(* IEC 61131-3 sources: plcassist-cli/packages/volt-lsp-iec/test-corpus/bakon-nano/Device/Plc Logic/Application/Library Manager/L_MC1P_MotionControlBasic, 488 files *)

(* ---- L_MC1P_CONSTANTS.gvl ---- *)
VAR_GLOBAL
	GC_EPS : LREAL := 1E-10;
	GC_EPS_REAL : LREAL := 1E-06;
	GC_WUPDATEFILTER : WORD := 10;
	GC_WINSTANCENCHAR : WORD := 100;
	GC_WTRACEMAX : WORD := 100;
	GC_IMPLIZITCALLS : INT := 100;
	GC_MAXRETAINAXIS : INT := 256;
	GC_MAXAXISCOUNT : INT := 256;
	GC_ENCFILTERCYCLESMAX : INT := 100;
	GC_DWCHECKIDTAPPETREF : DWORD := 16#DC34;
	GC_SQRT2 : LREAL := 1.4142135623730951;
	GC_PI : LREAL := 3.1415926535897931;
	GC_REC_STATE : LWORD := SHL(1, 0);
	GC_REC_OPMODE : LWORD := SHL(1, 1);
	GC_REC_POS : LWORD := SHL(1, 2);
	GC_REC_VEL : LWORD := SHL(1, 3);
	GC_REC_TORQUE : LWORD := SHL(1, 4);
	GC_REC_ERRORID : LWORD := SHL(1, 5);
	GC_REC_FOLLERROR : LWORD := SHL(1, 6);
	GC_REC_STATELENZE : LWORD := SHL(1, 7);
	GC_REC_STATELENZE2 : LWORD := SHL(1, 8);
	GC_REC_TPSTATE1 : LWORD := SHL(1, 9);
	GC_REC_TP1POS : LWORD := SHL(1, 10);
	GC_REC_TP1NEG : LWORD := SHL(1, 11);
	GC_REC_TP2POS : LWORD := SHL(1, 12);
	GC_REC_TP2NEG : LWORD := SHL(1, 13);
	GC_REC_DIGIN : LWORD := SHL(1, 14);
	GC_REC_STATESM : LWORD := SHL(1, 15);
	GC_REC_VLACTVELOCITY : LWORD := SHL(1, 16);
	GC_REC_ENCPOS : LWORD := SHL(1, 17);
	GC_REC_ENCVEL : LWORD := SHL(1, 18);
	GC_REC_TP1POSTIME : LWORD := SHL(1, 19);
	GC_REC_TP1NEGTIME : LWORD := SHL(1, 20);
	GC_REC_TP2POSTIME : LWORD := SHL(1, 21);
	GC_REC_TP2NEGTIME : LWORD := SHL(1, 22);
	GC_REC_TPSTATE2 : LWORD := SHL(1, 23);
	GC_REC_TP3POS : LWORD := SHL(1, 24);
	GC_REC_TP3NEG : LWORD := SHL(1, 25);
	GC_REC_TP4POS : LWORD := SHL(1, 26);
	GC_REC_TP4NEG : LWORD := SHL(1, 27);
	GC_REC_TP3POSTIME : LWORD := SHL(1, 28);
	GC_REC_TP3NEGTIME : LWORD := SHL(1, 29);
	GC_REC_TP4POSTIME : LWORD := SHL(1, 30);
	GC_REC_TP4NEGTIME : LWORD := SHL(1, 31);
	GC_REC_SAFETYCTRL : LWORD := SHL(1, 32);
	GC_REC_SAFETYSTATE : LWORD := SHL(1, 33);
	GC_REC_SAFETYIOSTATE : LWORD := SHL(1, 34);
	GC_REC_ENCPOSTIMESTAMP : LWORD := SHL(1, 35);
	GC_REC_STATELENZEEXT : LWORD := SHL(1, 36);
	GC_REC_SPEEDERROR : LWORD := SHL(1, 37);
	GC_REC_POSVALUE1616 : LWORD := SHL(1, 38);
	GC_REC_CONTROLEFFORT : LWORD := SHL(1, 39);
	GC_REC_ACTPOSMOTORCIA402ADV : LWORD := SHL(1, 40);
	GC_REC_TEXTREFID : LWORD := SHL(1, 41);
	GC_REC_POSTIMESTAMP : LWORD := SHL(1, 42);
	GC_REC_MAXDATAINDEX : WORD := 43;
	GC_TRANS_CTRL : LWORD := SHL(1, 0);
	GC_TRANS_OPMODE : LWORD := SHL(1, 1);
	GC_TRANS_POS : LWORD := SHL(1, 2);
	GC_TRANS_VEL : LWORD := SHL(1, 3);
	GC_TRANS_TORQUE : LWORD := SHL(1, 4);
	GC_TRANS_TORQUELIMPOS : LWORD := SHL(1, 5);
	GC_TRANS_TORQUELIMNEG : LWORD := SHL(1, 6);
	GC_TRANS_SPEEDLIMUP : LWORD := SHL(1, 7);
	GC_TRANS_SPEEDLIMLOW : LWORD := SHL(1, 8);
	GC_TRANS_TPCTRL1 : LWORD := SHL(1, 9);
	GC_TRANS_POSOFFSET : LWORD := SHL(1, 10);
	GC_TRANS_VELOFFSET : LWORD := SHL(1, 11);
	GC_TRANS_TORQUEOFFSET : LWORD := SHL(1, 12);
	GC_TRANS_SPEEDCTRLINT : LWORD := SHL(1, 13);
	GC_TRANS_CTRLLENZE : LWORD := SHL(1, 14);
	GC_TRANS_VLTARGETVELOCITY : LWORD := SHL(1, 16);
	GC_TRANS_BRKOVRD : LWORD := SHL(1, 17);
	GC_TRANS_CTRLLENZE2 : LWORD := SHL(1, 18);
	GC_TRANS_CTRLLENZE3 : LWORD := SHL(1, 19);
	GC_TRANS_CTRLLENZE4 : LWORD := SHL(1, 20);
	GC_TRANS_TPCTRL2 : LWORD := SHL(1, 21);
	GC_TRANS_SAFEPOS : LWORD := SHL(1, 22);
	GC_TRANS_SAFEPOSSTATUS : LWORD := SHL(1, 23);
	GC_TRANS_SPEEDLIMITSLS : LWORD := SHL(1, 24);
	GC_TRANS_MAXDATAINDEX : WORD := 25;
	NODATAMEMORYAVAILABLE : WORD := WORD#16#1;
	MEMORYINVALID : WORD := WORD#16#2;
	MEMORYNOTINITIALIZED : WORD := WORD#16#4;
	NODATAAVAILABLE : WORD := WORD#16#8;
	NOMEMORYAVAILABLEFORAXIS : WORD := WORD#16#10;
	NOMEMORYINAXISARRAY : WORD := WORD#16#20;
	AXISGUIDCHANGED : WORD := WORD#16#40;
	C_SERIALNUMBER : UINT := 3;
	C_MANUFACTURER : UINT := 5;
	C_SOFTWAREREVISION : UINT := 9;
	C_HARDWAREREVISION : UINT := 10;
	C_DEVICECLASS : UINT := 11;
	C_PRODUCTCODE : UINT := 13;
	C_UPDATE : UINT := 99;
	C_CONNECTORTYPEMOTIONAXISOLD : UINT := 1279;
	C_CONNECTORTYPEMOTIONAXIS : UINT := 34279;
	C_CONNECTORTYPEENCODERIOSLICE : UINT := 33024;
END_VAR

(* ---- L_MC1P_INTERNAL.gvl ---- *)
VAR_GLOBAL
	DWDUMMY : DWORD;
	XAPPFIRSTRUN : BOOL := FALSE;
	PANYCONNECTOR : POINTER TO IoConfigConnector;
	LMAXISRETAINHANDLING : L_MC1P_AxisRetainMangaement;
	DWTIMESTAMPSIMU : DWORD;
	XTIMESTAMPUPDATED : BOOL;
	LMAXISMGMT : L_MC1P_AxisManagementFunction;
	CDIENUMSTARTVALUE : DINT := 50000;
END_VAR

(* ---- L_MC1P_IAXIS_REF_BRAKE.itf ---- *)
INTERFACE L_MC1P_IAXIS_REF_BRAKE
END_INTERFACE

METHOD GETACTVALUESBRAKE
END_METHOD

METHOD SWITCHONCONTROL
VAR_INPUT
	XSWITCHONREQUEST : BOOL;
END_VAR
VAR_OUTPUT
	XSWITCHON : BOOL;
END_VAR
VAR_IN_OUT
	AXIS : AXIS_REF;
END_VAR
END_METHOD

METHOD SWITCHEDONSTATUS
VAR_INPUT
	XSWITCHEDONREQUEST : BOOL;
END_VAR
VAR_OUTPUT
	XSWITCHEDON : BOOL;
END_VAR
VAR_IN_OUT
	AXIS : AXIS_REF;
END_VAR
END_METHOD

(* ---- L_MC1P_IAXIS_REF_MASTERVALUES.itf ---- *)
INTERFACE L_MC1P_IAXIS_REF_MASTERVALUES
END_INTERFACE

METHOD GETDIRECTION : WORD
VAR_INPUT
	VALUESOURCE : MC_SOURCE;
END_VAR
END_METHOD

METHOD GETMASTERERROR : BOOL
VAR_OUTPUT
	EERRORID : L_IE1P_Error;
END_VAR
END_METHOD

METHOD GETSTEADYSTATE : POINTER TO L_MC1P_SteadyState
END_METHOD

(* ---- L_MC1P_IAXIS_REF_POOL.itf ---- *)
INTERFACE L_MC1P_IAXIS_REF_POOL
END_INTERFACE

METHOD GETAXISFROMPOOL : POINTER TO AXIS_REF
VAR_INPUT
	WINDEX : WORD;
END_VAR
END_METHOD

(* ---- L_MC1P_IAXISCOMMMAND.itf ---- *)
INTERFACE L_MC1P_IAXISCOMMMAND
END_INTERFACE

METHOD ABORTING
END_METHOD

METHOD CALCSTATUS
VAR_IN_OUT
	AXIS : _AXIS_REF_REAL;
END_VAR
END_METHOD

METHOD EXECUTE
END_METHOD

METHOD MAIN
END_METHOD

METHOD RESETCOMMANDERRORSTATE : BOOL
VAR_IN_OUT
	AXIS : _AXIS_REF_REAL;
END_VAR
END_METHOD

METHOD RESETSTATUSPARAMETER
END_METHOD

METHOD SETINCTANCEINFO
VAR_INPUT
	PSINSTANCENAME : POINTER TO STRING;
	ERRORITFID : DWORD;
END_VAR
END_METHOD

METHOD UPDATEAXISPOINTER
VAR_INPUT
	PAXIS : POINTER TO AXIS_REF;
END_VAR
END_METHOD

METHOD UPDATECOMMANDINTERFACE
VAR_IN_OUT
	CMD : USINT;
END_VAR
END_METHOD

(* ---- L_MC1P_IAXISCOMMMAND_AUTOTUNING.itf ---- *)
INTERFACE L_MC1P_IAXISCOMMMAND_AUTOTUNING
END_INTERFACE

METHOD CALCPROFILEPARAMS
VAR_IN_OUT
	AXIS : AXIS_REF;
END_VAR
END_METHOD

METHOD UPDATEPARAINTERFACE
VAR_IN_OUT
	SCPAR : L_MC1P_AutotuningPara;
END_VAR
END_METHOD

(* ---- L_MC1P_IAXISEXTENSION.itf ---- *)
INTERFACE L_MC1P_IAXISEXTENSION
END_INTERFACE

METHOD SETBASICINITIALISATION
VAR_INPUT
	ITFGENERICCONFIG : L_MC1P_IGenericAxisConfiguration;
END_VAR
VAR_IN_OUT
	AXIS : _AXIS_REF_REAL;
END_VAR
END_METHOD

(* ---- L_MC1P_IAXISSIMCALLSINGLESTEPS.itf ---- *)
INTERFACE L_MC1P_IAXISSIMCALLSINGLESTEPS
END_INTERFACE

METHOD SIMFINISH : BOOL
VAR_INPUT
	AXISID : INT;
	ITFMECHANICSIMULATION : L_MC1P_IMechanicSimulation;
END_VAR
VAR_IN_OUT
	AXIS : _AXIS_REF_REAL;
END_VAR
END_METHOD

METHOD SIMINSIDELOOP : BOOL
VAR_INPUT
	AXISID : INT;
	ISYSTEMSIMCOUNTER : INT;
	ITFMECHANICSIMULATION : L_MC1P_IMechanicSimulation;
END_VAR
END_METHOD

METHOD SIMPREPARE : BOOL
VAR_INPUT
	AXISID : INT;
	ITFMECHANICSIMULATION : L_MC1P_IMechanicSimulation;
END_VAR
VAR_IN_OUT
	AXIS : _AXIS_REF_REAL;
END_VAR
END_METHOD

(* ---- L_MC1P_IAXISSIMULATIONINTERFACE.itf ---- *)
INTERFACE L_MC1P_IAXISSIMULATIONINTERFACE
END_INTERFACE

METHOD ACTIVATESIMULATION
VAR_IN_OUT
	AXIS : _AXIS_REF_REAL;
END_VAR
END_METHOD

METHOD CALCULATEINPUTDATA
VAR_INPUT
	ITFKINSIM : L_MC1P_IKinematicSimulation;
END_VAR
VAR_IN_OUT
	AXIS : _AXIS_REF_REAL;
END_VAR
END_METHOD

METHOD CALCULATEOUTPUTDATA
VAR_INPUT
	ITFKINSIM : L_MC1P_IKinematicSimulation;
END_VAR
VAR_IN_OUT
	AXIS : _AXIS_REF_REAL;
END_VAR
END_METHOD

METHOD DISABLESIMULATION
VAR_IN_OUT
	AXIS : _AXIS_REF_REAL;
END_VAR
END_METHOD

(* ---- L_MC1P_ICOMMMUNICATIONSIMULATION.itf ---- *)
INTERFACE L_MC1P_ICOMMMUNICATIONSIMULATION
END_INTERFACE

METHOD GETCOMMSTATE : L_DCO_CommState
VAR_INPUT
	PAXISCOMM : POINTER TO _AXIS_REF_COM;
END_VAR
END_METHOD

METHOD PARREAD
VAR_INPUT
	WIDX : DWORD;
END_VAR
END_METHOD

METHOD PARREAD_GETOUTPUT
VAR_INPUT
	WIDX : DWORD;
END_VAR
VAR_OUTPUT
	SZDATAREAD : CAA_SIZE;
	XDONE : BOOL;
	XERROR : BOOL;
	WERROR : WORD;
END_VAR
END_METHOD

METHOD PARREAD_SETINPUT
VAR_INPUT
	WIDX : DWORD;
	XEXECUTE : BOOL;
	WINDEX : WORD;
	BYSUBINDEX : BYTE;
	PBUFFER : POINTER TO BYTE;
	SZSIZE : UDINT;
	UDITIMEOUT : UDINT;
	XSLOTB : BOOL;
END_VAR
END_METHOD

METHOD PARWRITE
VAR_INPUT
	WIDX : DWORD;
END_VAR
END_METHOD

METHOD PARWRITE_GETOUTPUT
VAR_INPUT
	WIDX : DWORD;
END_VAR
VAR_OUTPUT
	XDONE : BOOL;
	XERROR : BOOL;
	WERROR : WORD;
END_VAR
END_METHOD

METHOD PARWRITE_SETINPUT
VAR_INPUT
	WIDX : DWORD;
	XEXECUTE : BOOL;
	WINDEX : WORD;
	BYSUBINDEX : BYTE;
	PBUFFER : POINTER TO BYTE;
	SZSIZE : UDINT;
	UDITIMEOUT : UDINT;
	XSLOTB : BOOL;
END_VAR
END_METHOD

METHOD RESTARTMASTER
VAR_INPUT
	XEXECUTE : BOOL;
	PAXIS : POINTER TO _AXIS_REF_COM;
END_VAR
VAR_OUTPUT
	XDONE : BOOL;
	XERROR : BOOL;
	XBUSY : BOOL;
	DWERROR : DWORD;
END_VAR
END_METHOD

(* ---- L_MC1P_ICOMMUNICATION.itf ---- *)
INTERFACE L_MC1P_ICOMMUNICATION
END_INTERFACE

METHOD FORWARDERROR
VAR_INPUT
	XENABLE : BOOL;
	XWARNING : BOOL;
	XERROR : BOOL;
	WERRORID : WORD;
	WTEXTREFID : WORD;
	XRESETERROR : BOOL := FALSE;
	AXISMODULEHANDLER : L_IMHP_IModuleHandler;
END_VAR
END_METHOD

METHOD GETCOMMPARAMETER
VAR_INPUT
	PCONNECTOR : POINTER TO IoConfigConnector;
END_VAR
VAR_OUTPUT
	PSLAVECONNECTOR : POINTER TO IoStandard.IoConfigConnector;
	UINETID : UINT;
	UIDEVICEID : UINT;
	XSENDFRAMEATTASKSTART : BOOL;
	UDIPRODUCTCODE : DWORD;
	PMASTERCONNECTOR : POINTER TO IoStandard.IoConfigConnector;
END_VAR
END_METHOD

METHOD GETCOMMSTATE : L_DCO_CommState
VAR_INPUT
	PAXISCOMM : POINTER TO _AXIS_REF_COM;
END_VAR
END_METHOD

METHOD GETPDINEQPDOUT : BOOL
END_METHOD

METHOD PARREAD
VAR_INPUT
	WIDX : DWORD;
END_VAR
END_METHOD

METHOD PARREAD_GETOUTPUT
VAR_INPUT
	WIDX : DWORD;
END_VAR
VAR_OUTPUT
	SZDATAREAD : CAA_SIZE;
	XDONE : BOOL;
	XERROR : BOOL;
	WERROR : WORD;
END_VAR
END_METHOD

METHOD PARREAD_SETINPUT
VAR_INPUT
	WIDX : DWORD;
	XEXECUTE : BOOL;
	WINDEX : WORD;
	BYSUBINDEX : BYTE;
	PBUFFER : POINTER TO BYTE;
	SZSIZE : UDINT;
	UDITIMEOUT : UDINT;
END_VAR
END_METHOD

METHOD PARWRITE
VAR_INPUT
	WIDX : DWORD;
END_VAR
END_METHOD

METHOD PARWRITE_GETOUTPUT
VAR_INPUT
	WIDX : DWORD;
END_VAR
VAR_OUTPUT
	XDONE : BOOL;
	XERROR : BOOL;
	WERROR : WORD;
END_VAR
END_METHOD

METHOD PARWRITE_SETINPUT
VAR_INPUT
	WIDX : DWORD;
	XEXECUTE : BOOL;
	WINDEX : WORD;
	BYSUBINDEX : BYTE;
	PBUFFER : POINTER TO BYTE;
	SZSIZE : UDINT;
	UDITIMEOUT : UDINT;
END_VAR
END_METHOD

METHOD RESET
END_METHOD

METHOD RESTARTMASTER
VAR_INPUT
	XEXECUTE : BOOL;
	PAXIS : POINTER TO _AXIS_REF_COM;
END_VAR
VAR_OUTPUT
	XDONE : BOOL;
	XERROR : BOOL;
	XBUSY : BOOL;
	DWERROR : DWORD;
END_VAR
END_METHOD

METHOD SETBASICINITIALISATION
VAR_IN_OUT
	AXIS : _AXIS_REF_REAL;
END_VAR
END_METHOD

METHOD SETCOMPONENTINFO
VAR_INPUT
	DATASELECTION : WORD;
	SDATA : STRING;
END_VAR
END_METHOD

(* ---- L_MC1P_ICOMPENSATIONINTERFACE.itf ---- *)
INTERFACE L_MC1P_ICOMPENSATIONINTERFACE
END_INTERFACE

METHOD GETOFFSETVALUES
VAR_OUTPUT
	LROFFSETPOS : LREAL;
	LROFFSETVEL : LREAL;
	LROFFSETACC : LREAL;
END_VAR
END_METHOD

(* ---- L_MC1P_ICONFIGUREDRIVE.itf ---- *)
INTERFACE L_MC1P_ICONFIGUREDRIVE
END_INTERFACE

METHOD DOFUNCTION : BOOL
VAR_INPUT
	XEXECUTE : BOOL;
	WOFFSET : WORD;
END_VAR
VAR_OUTPUT
	XDONE : BOOL;
	XERROR : BOOL;
	XBUSY : BOOL;
	EERRORID : WORD;
END_VAR
VAR_IN_OUT
	AXIS : _AXIS_REF_REAL;
END_VAR
END_METHOD

METHOD GETADDITIONALCONFIGINFO : POINTER TO L_MC1P_AdditionalConfigInfo
END_METHOD

METHOD GETINSTANCE : POINTER TO BYTE
END_METHOD

METHOD RESET : BOOL
END_METHOD

(* ---- L_MC1P_ICONTROLLERADAPTION.itf ---- *)
INTERFACE L_MC1P_ICONTROLLERADAPTION
END_INTERFACE

METHOD CALCADAPTIONCURVE : LREAL
VAR_INPUT
	LRSETVEL : LREAL;
END_VAR
VAR_IN_OUT
	AXIS : _AXIS_REF_REAL;
END_VAR
END_METHOD

(* ---- L_MC1P_ICONTROLLERINTERFACE.itf ---- *)
INTERFACE L_MC1P_ICONTROLLERINTERFACE
END_INTERFACE

METHOD CALCCONTROLLER
VAR_INPUT
	LRSETPOSITION : LREAL;
	LRSETVELOCITY : LREAL;
	LRSETACCELERATION : LREAL;
	LRSETTORQUE : LREAL;
	LRSETJERK : LREAL;
	LRACTPOSITIONIN : LREAL;
	LRACTVELOCITYIN : LREAL;
	LRACTACCELERATIONIN : LREAL;
	LRACTTORQUEIN : LREAL;
END_VAR
VAR_OUTPUT
	LRSETPOSITIONOUT : LREAL;
	LRSETVELOCITYOUT : LREAL;
	LRSETACCELERATIONOUT : LREAL;
	LRSETTORQUEOUT : LREAL;
END_VAR
VAR_IN_OUT
	AXIS : _AXIS_REF_REAL;
END_VAR
END_METHOD

(* ---- L_MC1P_IDRIVESCALING.itf ---- *)
INTERFACE L_MC1P_IDRIVESCALING
END_INTERFACE

METHOD CALCACCFACTOR : BOOL
VAR_OUTPUT
	LRSCALEUNITTOACC : LREAL;
	LRSCALEACCTOUNIT : LREAL;
END_VAR
VAR_IN_OUT
	AXIS : _AXIS_REF_REAL;
END_VAR
END_METHOD

METHOD CALCSPEEDFACTOR : BOOL
VAR_OUTPUT
	LRSCALEUNITTOSPEED : LREAL;
	LRSCALESPEEDTOUNIT : LREAL;
END_VAR
VAR_IN_OUT
	AXIS : _AXIS_REF_REAL;
END_VAR
END_METHOD

METHOD CALCTORQUEFACTOR : BOOL
VAR_OUTPUT
	LRSCALETORQUETONORM : LREAL;
	LRSCALETORQUETONORM2 : LREAL;
	LRSCALENORMTOTORQUE : LREAL;
END_VAR
VAR_IN_OUT
	AXIS : _AXIS_REF_REAL;
END_VAR
END_METHOD

METHOD CHECKVALIDPOSRESOLUTION : BOOL
VAR_INPUT
	DWPOSRESOLUTION : DWORD;
END_VAR
END_METHOD

METHOD GETDEFAULTTORQUE : LREAL
VAR_INPUT
	LRREFTORQUE : LREAL;
END_VAR
END_METHOD

METHOD POSDIFFTOSPEEDINC : DINT
VAR_INPUT
	DIPOSDIFF : DINT := 0;
	DWFACTOR : DWORD := 1000;
END_VAR
VAR_IN_OUT
	AXIS : _AXIS_REF_REAL;
END_VAR
END_METHOD

METHOD SPEEDTOPOSDIFFINC : DINT
VAR_INPUT
	DISPEED : DINT := 0;
	DWFACTOR : DWORD := 1000;
END_VAR
VAR_IN_OUT
	AXIS : _AXIS_REF_REAL;
	DIRES : DINT;
END_VAR
END_METHOD

(* ---- L_MC1P_IDRIVESPECIFICIMPLBASE.itf ---- *)
INTERFACE L_MC1P_IDRIVESPECIFICIMPLBASE
END_INTERFACE

METHOD CALCAFTERREADINPUTS
VAR_IN_OUT
	AXIS : _AXIS_REF_REAL;
END_VAR
END_METHOD

METHOD CALCBEFOREREADINPUTS
VAR_IN_OUT
	AXIS : _AXIS_REF_REAL;
END_VAR
END_METHOD

METHOD CALCBEFOREWRITEOUTPUTS
VAR_IN_OUT
	AXIS : _AXIS_REF_REAL;
END_VAR
END_METHOD

METHOD CHECKAVAILABLECONTROLMODE : BOOL
VAR_IN_OUT
	AXIS : _AXIS_REF_REAL;
	POSCTRLDRIVEAVAILABLE : L_IE1P_Error;
	POSCTRLPLCAVAILABLE : L_IE1P_Error;
	SPEEDCTRLDRIVEAVAILABLE : L_IE1P_Error;
	TORQUECTRLDRIVE : L_IE1P_Error;
END_VAR
END_METHOD

METHOD CHECKRESETHOMEPOS
VAR_INPUT
	WFDBSTATUSWORD : WORD;
END_VAR
VAR_IN_OUT
	AXIS : _AXIS_REF_REAL;
END_VAR
END_METHOD

METHOD CHECKSAFETYOPTIONAVAILABLE : BOOL
VAR_INPUT
	DWPRODUCTCODE : DWORD;
END_VAR
END_METHOD

METHOD COLLECTDRIVESTATE : BOOL
VAR_IN_OUT
	AXIS : _AXIS_REF_REAL;
	SCSTATEINFO : L_MC1P_DriveStateCollection;
END_VAR
END_METHOD

METHOD CONTROLDRIVE : BOOL
VAR_INPUT
	XENABLE : BOOL;
END_VAR
VAR_IN_OUT
	AXIS : _AXIS_REF_REAL;
END_VAR
END_METHOD

METHOD DRIVECONFIGDATA
VAR_INPUT
	PCONFIGINFO : POINTER TO L_MC1P_AdditionalConfigInfo;
END_VAR
VAR_IN_OUT
	AXIS : _AXIS_REF_REAL;
END_VAR
END_METHOD

METHOD DRIVEFAULTSTATUS : BOOL
VAR_IN_OUT
	AXIS : _AXIS_REF_REAL;
	SCSTATEINFO : L_MC1P_DriveStateCollection;
END_VAR
END_METHOD

METHOD GETBRAKE : POINTER TO L_MC1P_BrakeControlBase
VAR_IN_OUT
	AXIS : _AXIS_REF_REAL;
END_VAR
END_METHOD

METHOD GETBRAKESERVICE : POINTER TO L_MC1P_BrakeService
VAR_IN_OUT
	AXIS : _AXIS_REF_REAL;
END_VAR
END_METHOD

METHOD GETCAUSEOFCINH : WORD
VAR_IN_OUT
	AXIS : _AXIS_REF_REAL;
END_VAR
END_METHOD

METHOD GETFDBSTATUSWORD : WORD
VAR_IN_OUT
	AXIS : _AXIS_REF_REAL;
END_VAR
END_METHOD

METHOD GETIECADRESS : BOOL
VAR_IN_OUT
	AXIS : _AXIS_REF_REAL;
	M_PPDOINFOCONNECTOR : POINTER TO IoConfigConnector;
	ATRANSELEMENT : ARRAY [1.._AXIS_REF_REAL.c_wMaxTransElem] OF L_MC1P_MappedElement;
	WTRANSELEMENTS : WORD;
	LWTRANSDATA : LWORD;
	LWRECDATA : LWORD;
	WRECEIVEELEMENTS : WORD;
	ARECEIVEELEMENT : ARRAY [1.._AXIS_REF_REAL.c_wMaxRecElem] OF L_MC1P_MappedElement;
END_VAR
END_METHOD

METHOD GETOPTIONALACTVEL : BOOL
VAR_IN_OUT
	LRVEL : LREAL;
END_VAR
END_METHOD

METHOD GETRECEIVEDATAIMPL : DWORD
VAR_INPUT
	LWMASK : LWORD;
END_VAR
VAR_IN_OUT
	AXIS : _AXIS_REF_REAL;
END_VAR
END_METHOD

METHOD GETSTATUSWORDS
VAR_OUTPUT
	STATUSWORD1 : WORD;
	STATUSWORD2 : WORD;
	STATUSWORD3 : WORD;
	STATUSWORD4 : WORD;
END_VAR
VAR_IN_OUT
	AXIS : _AXIS_REF_REAL;
END_VAR
END_METHOD

METHOD GETTRANSMITDATAIMPL : DWORD
VAR_INPUT
	LWMASK : LWORD;
END_VAR
VAR_IN_OUT
	AXIS : _AXIS_REF_REAL;
END_VAR
END_METHOD

METHOD GETTRANSMITDATALREALIMPL : LREAL
VAR_INPUT
	LWMASK : LWORD;
END_VAR
VAR_IN_OUT
	AXIS : _AXIS_REF_REAL;
END_VAR
END_METHOD

METHOD HOMECONFIG : BOOL
VAR_INPUT
	LRPOSITION : LREAL;
END_VAR
VAR_OUTPUT
	WINDEX : WORD;
	BYSUBINDEX : BYTE;
	BYNROFBYTE : BYTE;
	DWDATA : DWORD;
	XWRITEPARAM : BOOL;
	XDONE : BOOL;
	XERROR : BOOL;
END_VAR
VAR_IN_OUT
	AXIS : _AXIS_REF_REAL;
	SCHOMEDATA : L_MC1P_HomeParameter;
	WSTEP : WORD;
END_VAR
END_METHOD

METHOD HOMEPOSPERMANENTSETACTIVE : BOOL
VAR_IN_OUT
	AXIS : _AXIS_REF_REAL;
END_VAR
END_METHOD

METHOD RECEIVEPARAMETER
VAR_INPUT
	WPARAMETER : WORD;
	PADRESS : POINTER TO BYTE;
	WSIZE : WORD;
END_VAR
VAR_IN_OUT
	AXIS : _AXIS_REF_REAL;
END_VAR
END_METHOD

METHOD RECEIVEPARAMETERCALC
VAR_IN_OUT
	AXIS : _AXIS_REF_REAL;
	DATA : ARRAY [1..L_MC1P_Constants.gc_Rec_MaxDataIndex] OF POINTER TO L_MC1P_MappedElement;
END_VAR
END_METHOD

METHOD RESETDRIVECONTROL
VAR_INPUT
	XRESETDRIVEERROR : BOOL;
END_VAR
END_METHOD

METHOD RESTOREADDITIONALRETAINDATA
VAR_INPUT
	PDATA : POINTER TO L_MC1P_uRetainData;
END_VAR
END_METHOD

METHOD SETAXISPROPERTIES
VAR_IN_OUT
	AXIS : _AXIS_REF_REAL;
	AXISPROPERTIES : L_MC1P_AxisProperties;
END_VAR
END_METHOD

METHOD SETAXISSTATUSWORD
VAR_IN_OUT
	AXIS : _AXIS_REF_REAL;
	DWAXISSTATUS : DWORD;
END_VAR
END_METHOD

METHOD SETBASICINITIALISATION
VAR_IN_OUT
	AXIS : _AXIS_REF_REAL;
END_VAR
END_METHOD

METHOD SETCONTROLWORDS
VAR_INPUT
	CONTROLWORD1 : WORD;
	CONTROLWORD2 : WORD;
	CONTROLWORD3 : WORD;
	CONTROLWORD4 : WORD;
END_VAR
VAR_IN_OUT
	AXIS : _AXIS_REF_REAL;
END_VAR
END_METHOD

METHOD SETDCBRAKE
VAR_INPUT
	XSETDCBRAKE : BOOL;
END_VAR
VAR_OUTPUT
	XDCBRAKEACTIVE : BOOL;
END_VAR
VAR_IN_OUT
	AXIS : _AXIS_REF_REAL;
END_VAR
END_METHOD

METHOD SETDRIVECONFIGINIT
VAR_IN_OUT
	AXIS : _AXIS_REF_REAL;
END_VAR
END_METHOD

METHOD SETSPEEDCTRLLIMITATION : BOOL
VAR_INPUT
	XLIMIT : BOOL;
END_VAR
VAR_IN_OUT
	AXIS : _AXIS_REF_REAL;
END_VAR
END_METHOD

METHOD SETSPEEDCTRLLOADVALUE
VAR_INPUT
	XLOAD : BOOL;
	LRVALUE : LREAL;
END_VAR
VAR_IN_OUT
	AXIS : _AXIS_REF_REAL;
END_VAR
END_METHOD

METHOD STOREADDITIONALRETAINDATA
VAR_INPUT
	PDATA : POINTER TO L_MC1P_uRetainData;
END_VAR
END_METHOD

METHOD TRANSMITPARAMETER
VAR_INPUT
	WPARAMETER : WORD;
	PADRESS : POINTER TO BYTE;
	WSIZE : WORD;
END_VAR
VAR_IN_OUT
	AXIS : _AXIS_REF_REAL;
END_VAR
END_METHOD

METHOD TRANSMITPARAMETERCALC
VAR_IN_OUT
	AXIS : _AXIS_REF_REAL;
	DATA : ARRAY [1..L_MC1P_Constants.gc_Trans_MaxDataIndex] OF POINTER TO L_MC1P_MappedElement;
END_VAR
END_METHOD

METHOD UPDATEMAPPING
VAR_INPUT
	PTASKMAPLIST : POINTER TO IoStandard.IoConfigTaskMap;
	NCOUNT : DINT;
	PPDOINFOCONNECTOR : POINTER TO IoConfigConnector;
END_VAR
VAR_IN_OUT
	AXIS : _AXIS_REF_REAL;
END_VAR
END_METHOD

(* ---- L_MC1P_IDRIVEUTILS.itf ---- *)
INTERFACE L_MC1P_IDRIVEUTILS
END_INTERFACE

METHOD ACTIVATEAPPCREDITS
VAR_INPUT
	XACTIVATE : BOOL;
END_VAR
END_METHOD

METHOD GETMULTIAXISINFO
VAR_IN_OUT
	MULTIAXISINFO : L_MC1P_MultiAxisInfo;
END_VAR
END_METHOD

METHOD GETRETAINMEMINFO : L_MC1P_RetainDataType
VAR_OUTPUT
	MEMINFO : L_MC1P_uAxisRetainInfo;
END_VAR
END_METHOD

METHOD RESETCONNECTION : L_IE1P_Error
VAR_INPUT
	ITFCALLEDFUNCITON : L_IF1P_IFunctionConnection;
	EDISCONNECTMODE : L_IF1P_DisconnectMode;
	XDISCONNECTEXISTINGCONNECTION : BOOL;
END_VAR
END_METHOD

METHOD SETCONNECTION
VAR_INPUT
	AXISCONNECTION : L_IF1P_IFunctionConnection;
END_VAR
END_METHOD

(* ---- L_MC1P_IENCODERINTERFACE.itf ---- *)
INTERFACE L_MC1P_IENCODERINTERFACE
END_INTERFACE

METHOD ENCNEWHOMEPOSLOADED : BOOL
VAR_INPUT
	DWCALLYCLE : DWORD;
	DWDELAY : DWORD;
END_VAR
END_METHOD

METHOD ENCRESETACTPOS
END_METHOD

METHOD ENCRESETHOMEPOS
VAR_INPUT
	ERESETINFO : L_IE1P_Error;
END_VAR
END_METHOD

METHOD ENCSETHOMEPOSITION
VAR_INPUT
	POSITION : LREAL;
	RELATIVE : BOOL;
	POSDIFF : LREAL;
	EHOMEPOSINFO : L_IE1P_Error;
END_VAR
END_METHOD

METHOD ENCSIGNALVALID : BOOL
VAR_OUTPUT
	XSIGNALVALIDOLD : BOOL;
	EENCERRORID : L_IE1P_Error;
END_VAR
END_METHOD

METHOD GETACTPOSINCR : DINT
END_METHOD

METHOD GETACTPOSINCR1616 : DINT
END_METHOD

METHOD GETACTVALUES
VAR_OUTPUT
	LRACTPOS : LREAL;
	LRACTVEL : LREAL;
	LRACTACC : LREAL;
	LRACTPOSUNFILTERED : LREAL;
	LRACTPOSROUNDS : LREAL;
END_VAR
END_METHOD

METHOD GETAXISINSTANCE : POINTER TO _AXIS_REF_REAL
END_METHOD

METHOD GETCONFIGCHANGED : BOOL
END_METHOD

METHOD GETHOMEPOSAVAILABLE : BOOL
END_METHOD

METHOD SETHOMEPOSAVAILABLE
VAR_INPUT
	XHOMEPOSAVAILABLE : BOOL;
END_VAR
END_METHOD

(* ---- L_MC1P_IENCODERPOSFILTER.itf ---- *)
INTERFACE L_MC1P_IENCODERPOSFILTER
END_INTERFACE

METHOD CALCULATE
VAR_INPUT
	LRCYCPOSIN : LREAL;
	LRCYCVELIN : LREAL;
END_VAR
VAR_OUTPUT
	LRCYCPOSOUT : LREAL;
	LRCYCVELOUT : LREAL;
	WFILTERSTATE : WORD;
END_VAR
END_METHOD

METHOD INIT
END_METHOD

METHOD RESET
END_METHOD

(* ---- L_MC1P_IERRORHANDLINGAXISSYSTEMS.itf ---- *)
INTERFACE L_MC1P_IERRORHANDLINGAXISSYSTEMS
END_INTERFACE

METHOD CLEARERRORINAXISSYSTEM
VAR_INPUT
	INSTANCEID : DWORD := 0;
END_VAR
END_METHOD

METHOD GETERRORITFID : DWORD
END_METHOD

METHOD NOTIFYERRORINAXISSYSTEM : BOOL
VAR_INPUT
	WERRORID : L_IE1P_Error := 0;
	INSTANCEID : DWORD := 0;
	PSINSTANCENAME : POINTER TO BYTE := 0;
	EERRORREACTION : L_IE1P_SeverityLevel := 0;
END_VAR
END_METHOD

(* ---- L_MC1P_IEXTENDEDMAPPINGACCESS.itf ---- *)
INTERFACE L_MC1P_IEXTENDEDMAPPINGACCESS
END_INTERFACE

METHOD GETIECADRESS
VAR_INPUT
	AXISCONNECTOR : POINTER TO IoConfigConnector;
END_VAR
END_METHOD

METHOD GETMAPPEDDATA : POINTER TO BYTE
VAR_INPUT
	UIINDEX : WORD;
	USISUBINDEX : USINT;
	USISIZE : USINT;
	XWRITEACCESS : BOOL;
	PADDDATA : POINTER TO BYTE;
	PXWAITFORINITACCESS : POINTER TO BOOL;
END_VAR
VAR_OUTPUT
	EERRORID : L_IE1P_Error;
	XERROR : BOOL;
	USISIZEACT : USINT;
END_VAR
END_METHOD

METHOD GETMAPPEDDATASUPPORT : BOOL
END_METHOD

METHOD RESETOUTPUTMAPPINGOBJECTS : BOOL
END_METHOD

(* ---- L_MC1P_IGENERICAXISCONFIGURATION.itf ---- *)
INTERFACE L_MC1P_IGENERICAXISCONFIGURATION
END_INTERFACE

METHOD CALCAFTERREADINPUTS
VAR_IN_OUT
	AXIS : _AXIS_REF_REAL;
	DRIVESPECIFIC : L_MC1P_DriveSpecific_Generic;
END_VAR
END_METHOD

METHOD CALCBEFOREREADINPUTS
VAR_IN_OUT
	AXIS : _AXIS_REF_REAL;
	DRIVESPECIFIC : L_MC1P_DriveSpecific_Generic;
END_VAR
END_METHOD

METHOD CALCBEFOREWRITEOUTPUTS
VAR_IN_OUT
	AXIS : _AXIS_REF_REAL;
	DRIVESPECIFIC : L_MC1P_DriveSpecific_Generic;
END_VAR
END_METHOD

METHOD DRIVECONFIG
VAR_INPUT
	WOFFSET : WORD;
END_VAR
VAR_OUTPUT
	XCONFIGBUSY : BOOL;
	XWAITFORPARAMETERWRITEDONE : BOOL;
	XWAITFORPARAMETERREADDONE : BOOL;
	XREADSTRING : BOOL;
	DWWRITEDATA : DWORD;
	WINDEX : WORD;
	BYSUBINDEX : BYTE;
	BYNROFBYTE : BYTE;
END_VAR
VAR_IN_OUT
	AXIS : _AXIS_REF_REAL;
	CONFIGINFO : L_MC1P_AdditionalConfigInfo;
	WSTEP : WORD;
	EERRORID : WORD;
	DWREADDATA : DWORD;
	SREADDATA : STRING(255);
END_VAR
END_METHOD

METHOD GETADDITIONALSTATEINFOS : BOOL
VAR_IN_OUT
	AXIS : _AXIS_REF_REAL;
	DRIVESPECIFIC : L_MC1P_DriveSpecific_Generic;
	SCSTATEINFO : L_MC1P_DriveStateCollection;
END_VAR
END_METHOD

METHOD GETHOMINGSTATE
VAR_INPUT
	WHOMESTATE : WORD;
END_VAR
VAR_IN_OUT
	AXIS : _AXIS_REF_REAL;
	XHOMEPOSAVAILABLEDRIVE : BOOL;
END_VAR
END_METHOD

METHOD HOMECONFIG
VAR_INPUT
	LRPOSITION : LREAL;
END_VAR
VAR_OUTPUT
	XCONFIGBUSY : BOOL;
	XERROR : BOOL;
	WINDEX : WORD;
	BYSUBINDEX : BYTE;
	BYNROFBYTE : BYTE;
	DWDATA : DWORD;
	XWRITEPARAM : BOOL;
END_VAR
VAR_IN_OUT
	AXIS : _AXIS_REF_REAL;
	SCHOMEDATA : L_MC1P_HomeParameter;
	WSTEP : WORD;
END_VAR
END_METHOD

METHOD RECEIVEPARAMETERCALC
VAR_IN_OUT
	AXIS : _AXIS_REF_REAL;
	DATA : ARRAY [1..L_MC1P_Constants.gc_Rec_MaxDataIndex] OF POINTER TO L_MC1P_MappedElement;
	DRIVESPECIFIC : L_MC1P_DriveSpecific_Generic;
END_VAR
END_METHOD

METHOD TRANSMITPARAMETERCALC
VAR_IN_OUT
	AXIS : _AXIS_REF_REAL;
	DATA : ARRAY [1..L_MC1P_Constants.gc_Trans_MaxDataIndex] OF POINTER TO L_MC1P_MappedElement;
	DRIVESPECIFIC : L_MC1P_DriveSpecific_Generic;
END_VAR
END_METHOD

(* ---- L_MC1P_IKINEMATICMASTER.itf ---- *)
INTERFACE L_MC1P_IKINEMATICMASTER
END_INTERFACE

METHOD ACTIVATEHOMESIGNALMONITORINGSLAVE
END_METHOD

METHOD ADDOFFSETVALUESFORMASTER
VAR_IN_OUT
	LRSETPOSITION : LREAL;
	LRSETVELOCITY : LREAL;
	LRSETACCELERATION : LREAL;
	LRSETTORQUE : LREAL;
END_VAR
END_METHOD

METHOD FINISHHOMINGFORMASTERAXIS : BOOL
END_METHOD

METHOD GETERRORACTIVEMAINAXIS : BOOL
END_METHOD

METHOD GETERRORSETVALUESFROMMAINAXIS : BOOL
VAR_INPUT
	XCONTROLLEDSTOPPOSSIBLE : BOOL;
END_VAR
VAR_OUTPUT
	XSETQSP : BOOL;
	XSETCINH : BOOL;
END_VAR
END_METHOD

METHOD GETMASTERAXISINSTANCE : POINTER TO AXIS_REF
END_METHOD

METHOD SETERRORMAINAXIS : BOOL
VAR_INPUT
	ESEVERITY : L_IE1P_SeverityLevel;
	WERRORID : WORD;
	DWEXTENDEDERRORINFO : DWORD;
END_VAR
END_METHOD

METHOD SWITCHROLE : BOOL
VAR_INPUT
	XSWITCH : BOOL;
END_VAR
END_METHOD

METHOD WAITHOMINGFORMASTERAXIS : BOOL
END_METHOD

METHOD FINISHBRAKETESTFORMASTERAXIS : BOOL
END_METHOD

METHOD FINISHGRINDINFORMASTERAXIS : BOOL
END_METHOD

METHOD WAITBRAKETESTFORMASTERAXIS : BOOL
END_METHOD

METHOD WAITGRINDINFORMASTERAXIS : BOOL
END_METHOD

(* ---- L_MC1P_IKINEMATICSIMULATION.itf ---- *)
INTERFACE L_MC1P_IKINEMATICSIMULATION
END_INTERFACE

METHOD CALLSYSSIM : BOOL
VAR_IN_OUT
	AXIS : _AXIS_REF_REAL;
END_VAR
END_METHOD

METHOD INITNEWCYCLE : BOOL
VAR_IN_OUT
	AXIS : _AXIS_REF_REAL;
END_VAR
END_METHOD

METHOD SETAXIS
VAR_INPUT
	AXISID : INT;
	PAXIS : POINTER TO _AXIS_REF_REAL;
END_VAR
END_METHOD

METHOD SETREQUIREDNUMBEROFAXIS
VAR_INPUT
	INUMAXIS : INT;
END_VAR
END_METHOD

(* ---- L_MC1P_IKINEMATICSLAVE.itf ---- *)
INTERFACE L_MC1P_IKINEMATICSLAVE
END_INTERFACE

METHOD ABORTHOMINGSLAVE : BOOL
END_METHOD

METHOD ACTIVATEHOMESIGNALMONITORINGMASTER
END_METHOD

METHOD ACTIVEMASTERHOMEPARAMETER
VAR_INPUT
	EHOMEMODE : L_MC1P_HomeMode;
	LRHOMEPOSITION : LREAL;
END_VAR
END_METHOD

METHOD ADDOFFSETVALUESFORSLAVE
VAR_IN_OUT
	LRSETPOSITION : LREAL;
	LRSETVELOCITY : LREAL;
	LRSETACCELERATION : LREAL;
	LRSETTORQUE : LREAL;
END_VAR
END_METHOD

METHOD CHECKHOMEPARAMETER : BOOL
VAR_OUTPUT
	XERROR : BOOL;
	EERRORID : L_IE1P_Error;
END_VAR
VAR_IN_OUT
	SCHOMEPARAMETER : L_MC1P_HomeParameter;
END_VAR
END_METHOD

METHOD DOHOMINGSLAVE : BOOL
END_METHOD

METHOD FINISHHOMINGFORSLAVEAXIS : BOOL
END_METHOD

METHOD GETERRORACTIVEFOLLOWAXIS : BOOL
END_METHOD

METHOD GETERRORSETVALUESFROMFOLLOWAXIS : BOOL
VAR_INPUT
	XCONTROLLEDSTOPPOSSIBLE : BOOL;
END_VAR
VAR_OUTPUT
	XSETQSP : BOOL;
	XSETCINH : BOOL;
END_VAR
END_METHOD

METHOD GETEXTERNALAUTOTUNINGITF : POINTER TO BYTE
VAR_INPUT
	XRESET : BOOL;
	UIACTUALATNBR : UINT;
END_VAR
VAR_OUTPUT
	WNBOFAUTOTUNINGS : WORD;
END_VAR
END_METHOD

METHOD GETMAXVEL : LREAL
VAR_IN_OUT
	LRVEL : LREAL;
END_VAR
END_METHOD

METHOD GETSETVALUESAVAILABLEMASTER : BOOL
END_METHOD

METHOD GETSLAVEAXISENABLED : BOOL
END_METHOD

METHOD GETSLAVEAXISHOMINGDONE : BOOL
END_METHOD

METHOD GETSLAVEAXISINSTANCE : POINTER TO AXIS_REF
END_METHOD

METHOD MOTIONALLOWED : BOOL
VAR_INPUT
	ETYPEFUNCTION : L_MC1P_TypeFunction;
END_VAR
VAR_OUTPUT
	EERRORCAUSE : L_IE1P_Error;
END_VAR
END_METHOD

METHOD RESETHOMEPOS
VAR_INPUT
	ERESETINFO : L_IE1P_Error;
	XRESETPOSITION : BOOL;
END_VAR
END_METHOD

METHOD RESTOREFOLLOWINGAXISERROR : BOOL
VAR_INPUT
	ESEVERITY : L_IE1P_SeverityLevel;
	WERRORID : WORD;
	DWEXTENDEDERRORINFO : DWORD;
END_VAR
END_METHOD

METHOD SETERRORFOLLOWAXIS : BOOL
VAR_INPUT
	ESEVERITY : L_IE1P_SeverityLevel;
	WERRORID : WORD;
	DWEXTENDEDERRORINFO : DWORD;
END_VAR
END_METHOD

METHOD SETHOMEPOS
VAR_INPUT
	POSITION : LREAL;
	RELATIVE : BOOL;
	XRESTARTPOSITIONING : BOOL := FALSE;
	EHOMEPOSINFO : L_IE1P_Error;
END_VAR
END_METHOD

METHOD SLAVEAXISRESETERROR : BOOL
END_METHOD

METHOD SLAVEAXISRESETPOSSIBLE : BOOL
END_METHOD

METHOD SWITCHROLE : BOOL
VAR_INPUT
	XSWITCH : BOOL;
END_VAR
END_METHOD

METHOD UPDATEABCSTATE : POINTER TO L_MC1P_AxisBasicControlOutput_Internal
END_METHOD

METHOD WAITHOMINGFORSLAVEAXIS : BOOL
END_METHOD

METHOD ABORTBRAKETESTSLAVE : BOOL
VAR_INPUT
	XMAINABORTED : BOOL;
END_VAR
END_METHOD

METHOD DOBRAKETESTSLAVE : BOOL
END_METHOD

METHOD FINISHBRAKETESTFORSLAVEAXIS : BOOL
END_METHOD

METHOD GETBTSTATUS : LREAL
END_METHOD

METHOD GETSLAVEAXISBRAKETESTDONE : BOOL
END_METHOD

METHOD WAITBRAKETESTFORSLAVEAXIS : BOOL
END_METHOD

METHOD ABORTGRINDINSLAVE : BOOL
VAR_INPUT
	XMAINABORTED : BOOL;
END_VAR
END_METHOD

METHOD DOGRINDINSLAVE : BOOL
END_METHOD

METHOD FINISHGRINDINFORSLAVEAXIS : BOOL
END_METHOD

METHOD GETACTIVEGRINDINCYCLESDONE : WORD
VAR_INPUT
	WCYCLESDONE : WORD;
END_VAR
END_METHOD

METHOD GETGICYCLES : LREAL
END_METHOD

METHOD GETGISTATUS : LREAL
END_METHOD

METHOD GETSLAVEAXISGRINDINDONE : BOOL
END_METHOD

METHOD WAITGRINDINFORSLAVEAXIS : BOOL
END_METHOD

(* ---- L_MC1P_ILMDATA.itf ---- *)
INTERFACE L_MC1P_ILMDATA
END_INTERFACE

METHOD ABORT : UDINT
END_METHOD

METHOD EXECUTE : UDINT
END_METHOD

(* ---- L_MC1P_IMANAGEMENTFUNCTION.itf ---- *)
INTERFACE L_MC1P_IMANAGEMENTFUNCTION
END_INTERFACE

METHOD COMPAREAXISNAME : BOOL
VAR_IN_OUT
	SAXISNAME : STRING;
END_VAR
END_METHOD

METHOD GETAXIS : POINTER TO AXIS_REF
END_METHOD

(* ---- L_MC1P_IMANIPULATEACTVALUES.itf ---- *)
INTERFACE L_MC1P_IMANIPULATEACTVALUES
END_INTERFACE

METHOD MANIPULATEACTVALUES
VAR_IN_OUT
	AXIS : AXIS_REF;
END_VAR
END_METHOD

(* ---- L_MC1P_IMANIPULATIONINTERFACE.itf ---- *)
INTERFACE L_MC1P_IMANIPULATIONINTERFACE
END_INTERFACE

METHOD CALCVALUES
VAR_INPUT
	XENABLE : BOOL;
	XRESET : BOOL;
	LRSETPOS : LREAL;
	LRSETVEL : LREAL;
	LRSETACC : LREAL;
	LRSETTORQUE : LREAL;
	XLOADPOSOFFSET : BOOL;
	LRPOSOFFSET : LREAL;
END_VAR
VAR_OUTPUT
	XACTIVE : BOOL;
	XERROR : BOOL;
	EERRORID : L_IE1P.L_IE1P_Error;
	LRSETPOSOUT : LREAL;
	LRSETVELOUT : LREAL;
	LRSETACCOUT : LREAL;
	LRSETTORQUEOUT : LREAL;
END_VAR
VAR_IN_OUT
	AXIS : Axis_REf;
END_VAR
END_METHOD

(* ---- L_MC1P_IMASTERINITINFO.itf ---- *)
INTERFACE L_MC1P_IMASTERINITINFO
END_INTERFACE

(* ---- L_MC1P_IMCPARAMETERACCESS.itf ---- *)
INTERFACE L_MC1P_IMCPARAMETERACCESS
END_INTERFACE

METHOD GETINSTANCEANDTYPE : BOOL
VAR_OUTPUT
	PINSTANCEPOINTER : POINTER TO BYTE;
	EAXISTYPE : L_MC1P_AxisType;
END_VAR
END_METHOD

METHOD HLP_GETPARAMETERPROPERTIES : BOOL
VAR_INPUT
	DIPARAMETER : DINT;
END_VAR
VAR_OUTPUT
	PPARAMADDR : POINTER TO BYTE;
	EORDINALTYPE : L_MC1P_OrdinalType;
	XREADWRITE : BOOL;
	LRUNITFACTOR : LREAL;
	LRDEFAULTVALUE : LREAL;
	WVALUERANGES : WORD;
	PVALUERANGES : POINTER TO L_MC1P_MinMaxValue;
END_VAR
END_METHOD

METHOD HLP_READBOOLPARAMETER : BOOL
VAR_INPUT
	PARAMETER : DINT;
	PXVALUE : POINTER TO BOOL;
END_VAR
END_METHOD

METHOD HLP_READPARAMETER : BOOL
VAR_INPUT
	PARAMETER : DINT;
	PLRVALUE : POINTER TO LREAL;
END_VAR
END_METHOD

METHOD HLP_WRITEBOOLPARAMETER : BOOL
VAR_INPUT
	PARAMETER : DINT;
	PXVALUE : POINTER TO BOOL;
END_VAR
VAR_OUTPUT
	WERRORID : WORD;
END_VAR
END_METHOD

METHOD HLP_WRITEPARAMETER : BOOL
VAR_INPUT
	PARAMETER : DINT;
	PLRVALUE : POINTER TO LREAL;
END_VAR
VAR_OUTPUT
	WERRORID : WORD;
END_VAR
END_METHOD

METHOD QUEUEDPARAMWRITINGACTIVE : BOOL
END_METHOD

(* ---- L_MC1P_IMECHANICSIMULATION.itf ---- *)
INTERFACE L_MC1P_IMECHANICSIMULATION
END_INTERFACE

METHOD CALLMECHANICSIMULATION : BOOL
VAR_INPUT
	AXISID : INT;
	XBRAKERELEASED : BOOL;
	LRACTTORQUE : LREAL;
	LRADDTORQUE : LREAL;
END_VAR
VAR_IN_OUT
	SCPARGENERAL : L_MC1P_ParGeneralMechanic;
END_VAR
END_METHOD

METHOD INITANDSCALEPARAMETER
VAR_INPUT
	AXISID : INT;
	LRTASKCYCLESYSSIM : LREAL;
	LRINVTASKCYCLESYSSIM : LREAL;
END_VAR
VAR_IN_OUT
	SCPARGENERAL : L_MC1P_ParGeneralMechanic;
END_VAR
END_METHOD

METHOD MECHANICSIMGETACTLOADVALUES
VAR_INPUT
	AXISID : INT;
END_VAR
VAR_OUTPUT
	LRACTLOADPOS : LREAL;
	LRACTLOADVEL : LREAL;
END_VAR
END_METHOD

METHOD MECHANICSIMGETACTVALUES
VAR_INPUT
	AXISID : INT;
END_VAR
VAR_OUTPUT
	LRACTPOS : LREAL;
	LRACTVEL : LREAL;
END_VAR
END_METHOD

METHOD SETLOADIDX
VAR_INPUT
	AXISID : INT;
	WIDXLOADMASS : WORD;
END_VAR
END_METHOD

METHOD SETSTARTPOSITION : BOOL
VAR_INPUT
	AXISID : INT;
	LRPOS : LREAL;
END_VAR
END_METHOD

(* ---- L_MC1P_IMOLACCESS.itf ---- *)
INTERFACE L_MC1P_IMOLACCESS
END_INTERFACE

METHOD SETMOLSTATES
VAR_INPUT
	WSETMOLSTATE : WORD := 0;
	WSETMOLMODE : WORD := 0;
END_VAR
END_METHOD

(* ---- L_MC1P_IPARA.itf ---- *)
INTERFACE L_MC1P_IPARA
END_INTERFACE

METHOD HLP_GETPARAMETERPROPERTIES : BOOL
VAR_INPUT
	PAXISREF : POINTER TO AXIS_REF;
	DIPARAMETER : DINT;
	XALLOWINVISIBLE : BOOL;
END_VAR
VAR_OUTPUT
	PPARAMADDR : POINTER TO BYTE;
	EORDINALTYPE : L_MC1P_OrdinalType;
	XREADWRITE : BOOL;
	LRUNITFACTOR : LREAL;
	LRDEFAULTVALUE : LREAL;
	WVALUERANGES : WORD;
	PVALUERANGES : POINTER TO L_MC1P_MinMaxValue;
END_VAR
END_METHOD

METHOD HLP_READBOOLPARAMETER : BOOL
VAR_INPUT
	PINPUTDATA : POINTER TO BYTE;
	PARAMETER : DINT;
	PXVALUE : POINTER TO BOOL;
	XALLOWINVISIBLE : BOOL;
END_VAR
END_METHOD

METHOD HLP_READPARAMETER : BOOL
VAR_INPUT
	PINPUTDATA : POINTER TO BYTE;
	PARAMETER : DINT;
	PLRVALUE : POINTER TO LREAL;
	XALLOWINVISIBLE : BOOL;
END_VAR
END_METHOD

METHOD HLP_WRITEBOOLPARAMETER : BOOL
VAR_INPUT
	PINPUTDATA : POINTER TO BYTE;
	PARAMETER : DINT;
	PXVALUE : POINTER TO BOOL;
	XALLOWINVISIBLE : BOOL;
END_VAR
VAR_OUTPUT
	WERRORID : WORD;
END_VAR
END_METHOD

METHOD HLP_WRITEPARAMETER : BOOL
VAR_INPUT
	PINPUTDATA : POINTER TO BYTE;
	PARAMETER : DINT;
	PLRVALUE : POINTER TO LREAL;
	XALLOWINVISIBLE : BOOL;
END_VAR
VAR_OUTPUT
	WERRORID : WORD;
END_VAR
END_METHOD

(* ---- L_MC1P_IPLIACCESS.itf ---- *)
INTERFACE L_MC1P_IPLIACCESS
END_INTERFACE

METHOD SETPPISTATES
VAR_INPUT
	WSETPPISTATE : WORD := 0;
	WSETPPIMODE : WORD := 0;
END_VAR
END_METHOD

(* ---- L_MC1P_IPOSPROFILECALCULATION.itf ---- *)
INTERFACE L_MC1P_IPOSPROFILECALCULATION
END_INTERFACE

METHOD CALCPROFILEDATA
VAR_INPUT
	PPOSPROFILERDATA : POINTER TO L_MC1P_PosProfiler;
	LRSTARTACC : LREAL;
	LRSTARTVEL : LREAL;
	LRSTARTPOS : LREAL;
	XVELMODE : BOOL;
END_VAR
VAR_OUTPUT
	XERROR : BOOL;
	DWSTATE : DWORD;
	DWPROFILETYPE : DWORD;
END_VAR
VAR_IN_OUT
	SCPROFILEDATA : L_MC1P_ProfileData;
	SCPROFILEPARAMETER : L_MC1P_ProfileParameter;
END_VAR
END_METHOD

METHOD PROFILEINTERPOLATOR : BOOL
VAR_INPUT
	PPOSPROFILERDATA : POINTER TO L_MC1P_PosProfiler;
	LREVALTIME : LREAL;
END_VAR
VAR_OUTPUT
	DWSTATE : DWORD;
	LRSETPOS : LREAL;
	LRSETVEL : LREAL;
	LRSETACC : LREAL;
END_VAR
VAR_IN_OUT
	SCPROFILEDATA : L_MC1P_ProfileData;
END_VAR
END_METHOD

METHOD STRETCHPROFILE
VAR_INPUT
	PPOSPROFILERDATA : POINTER TO L_MC1P_PosProfiler;
	LRTIMEBASE : LREAL;
END_VAR
VAR_IN_OUT
	SCPROFILEDATA : L_MC1P_ProfileData;
END_VAR
END_METHOD

(* ---- L_MC1P_IPOSPROFILERACTIVE.itf ---- *)
INTERFACE L_MC1P_IPOSPROFILERACTIVE
END_INTERFACE

(* ---- L_MC1P_IPOSSIGNALPROCESSING.itf ---- *)
INTERFACE L_MC1P_IPOSSIGNALPROCESSING
END_INTERFACE

METHOD CALCULATE : DINT
VAR_INPUT
	DIACTPOS : DINT;
	DWSAMPLETIME : DWORD;
	DWACTTIME : DWORD;
END_VAR
VAR_OUTPUT
	DIPOSOUT : DINT;
	XVELVALID : BOOL;
	DIVELOUT : DINT;
END_VAR
VAR_IN_OUT
	AXIS : _AXIS_REF_REAL;
END_VAR
END_METHOD

(* ---- L_MC1P_IRETAINFUNCTION.itf ---- *)
INTERFACE L_MC1P_IRETAINFUNCTION
END_INTERFACE

METHOD GETINITIALDATA : BOOL
VAR_INPUT
	PDATA : POINTER TO DWORD;
	INFO : DWORD;
END_VAR
END_METHOD

METHOD SETERRORINFO
VAR_INPUT
	WSTATE : WORD;
END_VAR
END_METHOD

METHOD SETINITIALDATA : BOOL
VAR_INPUT
	PDATA : POINTER TO DWORD;
END_VAR
END_METHOD

METHOD STOREDATA
VAR_INPUT
	PDATA : POINTER TO DWORD;
END_VAR
END_METHOD

(* ---- L_MC1P_IRETAINHANDLING.itf ---- *)
INTERFACE L_MC1P_IRETAINHANDLING
END_INTERFACE

METHOD GETINITIALRETAINDATA : POINTER TO L_MC1P_uRetainData
VAR_INPUT
	XNEWEST : BOOL;
END_VAR
END_METHOD

METHOD GETRETAINSTATE : WORD
VAR_OUTPUT
	WSTATERETAINERROR : WORD;
END_VAR
END_METHOD

METHOD REGISTERONRETAINDATAHANDLER
VAR_INPUT
	AXISGUID : L_MC1P_AxisGUID;
END_VAR
END_METHOD

METHOD RESET
END_METHOD

METHOD SETCONNECTEDGUID : BOOL
VAR_INPUT
	GUID : L_MC1P_AxisGUID;
END_VAR
END_METHOD

(* ---- L_MC1P_ISETSETVALUEMANIPULATORCUSTOM.itf ---- *)
INTERFACE L_MC1P_ISETSETVALUEMANIPULATORCUSTOM
END_INTERFACE

METHOD CALCULATE : L_IE1P_Error
VAR_INPUT
	UIINPUTDATAIDX : UINT;
	UIOUTPUTDATAIDX : UINT;
END_VAR
VAR_IN_OUT
	AXIS : AXIS_REF;
	LRSETPOS : LREAL;
	LRSETVEL : LREAL;
	LRSETACC : LREAL;
	LRSETTORQUE : LREAL;
END_VAR
END_METHOD

METHOD CALLCYCLIC : L_IE1P_Error
VAR_INPUT
	UIINPUTDATAIDX : UINT;
	UIOUTPUTDATAIDX : UINT;
END_VAR
VAR_IN_OUT
	AXIS : Axis_REf;
END_VAR
END_METHOD

METHOD CHECKINPUTDATA : L_IE1P_Error
VAR_INPUT
	UIINPUTDATAIDX : UINT;
	UIOUTPUTDATAIDX : UINT;
END_VAR
VAR_IN_OUT
	AXIS : AXIS_REF;
END_VAR
END_METHOD

METHOD ENABLEEXIT : L_IE1P_Error
VAR_INPUT
	UIINPUTDATAIDX : UINT;
	UIOUTPUTDATAIDX : UINT;
END_VAR
VAR_IN_OUT
	AXIS : AXIS_REF;
END_VAR
END_METHOD

METHOD ENABLEINIT : L_IE1P_Error
VAR_INPUT
	UIINPUTDATAIDX : UINT;
	UIOUTPUTDATAIDX : UINT;
END_VAR
VAR_IN_OUT
	AXIS : AXIS_REF;
END_VAR
END_METHOD

METHOD FREEZEINPUTPERCYCLE
VAR_INPUT
	UIINPUTDATAIDX : UINT;
END_VAR
END_METHOD

METHOD LOADOFFSET : L_IE1P_Error
VAR_INPUT
	UIINPUTDATAIDX : UINT;
	UIOUTPUTDATAIDX : UINT;
	OFFSET : LREAL;
END_VAR
VAR_IN_OUT
	AXIS : Axis_REf;
END_VAR
END_METHOD

METHOD PASSOUTPUTPERCYCLE
VAR_INPUT
	UIOUTPUTDATAIDX : UINT;
END_VAR
END_METHOD

METHOD READINPUTS : L_IE1P_Error
VAR_INPUT
	UIINPUTDATAIDX : UINT;
END_VAR
VAR_IN_OUT
	AXIS : Axis_REf;
END_VAR
END_METHOD

METHOD RESET : L_IE1P_Error
VAR_INPUT
	UIINPUTDATAIDX : UINT;
	UIOUTPUTDATAIDX : UINT;
END_VAR
VAR_IN_OUT
	AXIS : AXIS_REF;
END_VAR
END_METHOD

METHOD RESETOUTPUTS : L_IE1P_Error
VAR_INPUT
	UIOUTPUTDATAIDX : UINT;
END_VAR
VAR_IN_OUT
	AXIS : AXIS_REF;
END_VAR
END_METHOD

(* ---- L_MC1P_ISETVALUEMANIPULATIONINTERFACE.itf ---- *)
INTERFACE L_MC1P_ISETVALUEMANIPULATIONINTERFACE
END_INTERFACE

(* ---- L_MC1P_ITOUCHPROBEHANDLER.itf ---- *)
INTERFACE L_MC1P_ITOUCHPROBEHANDLER
END_INTERFACE

METHOD GETACTTPRECEIVEDATA : L_MC1P_TpReceiveData
END_METHOD

METHOD ISUPTODATE : BOOL
VAR_INPUT
	DWUPDATETIME : DWORD;
END_VAR
END_METHOD

METHOD RECDATAISVALID : BOOL
VAR_IN_OUT
	SCRECDATA : L_MC1P_TpReceiveData;
END_VAR
END_METHOD

(* ---- L_MC1P_ITPSOURCEAXIS.itf ---- *)
INTERFACE L_MC1P_ITPSOURCEAXIS
END_INTERFACE

METHOD GETPOINTERTOTPAXIS : POINTER TO _AXIS_REF_REAL
END_METHOD

(* ---- L_UBUP_ICALLORDERDEPENDENCY.itf ---- *)
INTERFACE L_UBUP_ICALLORDERDEPENDENCY
END_INTERFACE

METHOD CALC_OUTPUTS
END_METHOD

METHOD CALC_STATUSSIGNALS
END_METHOD

(* ---- GETBOOLEANPROPERTY.fun ---- *)
FUNCTION GETBOOLEANPROPERTY : BOOL
VAR_INPUT
	STKEY : WSTRING;
END_VAR
END_FUNCTION

(* ---- GETCOMPANY.fun ---- *)
FUNCTION GETCOMPANY : WSTRING
END_FUNCTION

(* ---- GETNUMBERPROPERTY.fun ---- *)
FUNCTION GETNUMBERPROPERTY : DINT
VAR_INPUT
	STKEY : WSTRING;
END_VAR
END_FUNCTION

(* ---- GETTEXTPROPERTY.fun ---- *)
FUNCTION GETTEXTPROPERTY : WSTRING
VAR_INPUT
	STKEY : WSTRING;
END_VAR
END_FUNCTION

(* ---- GETTEXTPROPERTY2.fun ---- *)
FUNCTION GETTEXTPROPERTY2 : POINTER TO WSTRING
VAR_INPUT
	STKEY : WSTRING;
END_VAR
END_FUNCTION

(* ---- GETTITLE.fun ---- *)
FUNCTION GETTITLE : WSTRING
END_FUNCTION

(* ---- GETVERSION.fun ---- *)
FUNCTION GETVERSION : VERSION
END_FUNCTION

(* ---- GETVERSIONPROPERTY.fun ---- *)
FUNCTION GETVERSIONPROPERTY : VERSION
VAR_INPUT
	STKEY : WSTRING;
END_VAR
END_FUNCTION

(* ---- L_MC1P_CHECKFORSENSORLESMODEIXXX.fun ---- *)
FUNCTION L_MC1P_CHECKFORSENSORLESMODEIXXX : BOOL
VAR_INPUT
	WMCTRLMODE : WORD;
END_VAR
END_FUNCTION

(* ---- L_MC1P_CODENUMBERTOPARAMETER.fun ---- *)
FUNCTION L_MC1P_CODENUMBERTOPARAMETER : DINT
VAR_INPUT
	DWCODENUMBER : DWORD;
	USISUBINDEX : USINT;
	UIBYTELENGTH : UINT;
END_VAR
END_FUNCTION

(* ---- L_MC1P_CODENUMBERTOPARAMETER2.fun ---- *)
FUNCTION L_MC1P_CODENUMBERTOPARAMETER2 : DINT
VAR_INPUT
	DWCODENUMBER : DWORD;
	USISUBINDEX : USINT;
	UIBYTELENGTH : UINT;
	XUNSIGNED : BOOL := FALSE;
END_VAR
END_FUNCTION

(* ---- L_MC1P_CONVERTPOSTOMODULOPOS.fun ---- *)
FUNCTION L_MC1P_CONVERTPOSTOMODULOPOS : LREAL
VAR_INPUT
	LRPOS : LREAL;
	LRPERIOD : LREAL;
END_VAR
END_FUNCTION

(* ---- L_MC1P_CONVERTPOSTOMODULOPOSEXTENDED.fun ---- *)
FUNCTION L_MC1P_CONVERTPOSTOMODULOPOSEXTENDED : LREAL
VAR_INPUT
	LRPOS : LREAL;
	LRPERIOD : LREAL;
END_VAR
END_FUNCTION

(* ---- L_MC1P_CONVERTPOSTOMODULOPOSFMOD.fun ---- *)
FUNCTION L_MC1P_CONVERTPOSTOMODULOPOSFMOD : LREAL
VAR_INPUT
	LRPOS : LREAL;
	LRPERIOD : LREAL;
END_VAR
END_FUNCTION

(* ---- L_MC1P_DIV.fun ---- *)
FUNCTION L_MC1P_DIV : LREAL
VAR_INPUT
	A : LREAL;
	B : LREAL;
END_VAR
END_FUNCTION

(* ---- L_MC1P_FINDDRIVECONNECTORFROMENCODER.fun ---- *)
FUNCTION L_MC1P_FINDDRIVECONNECTORFROMENCODER : POINTER TO IoConfigConnector
VAR_INPUT
	PCONNECTOR : POINTER TO IoConfigConnector;
END_VAR
END_FUNCTION

(* ---- L_MC1P_FINDOWNSLICEPOSITIONS131.fun ---- *)
FUNCTION L_MC1P_FINDOWNSLICEPOSITIONS131 : BOOL
VAR_INPUT
	M_PCONNECTOR : POINTER TO IoConfigConnector;
END_VAR
VAR_OUTPUT
	WSLICEPOSITION : WORD;
END_VAR
END_FUNCTION

(* ---- L_MC1P_FINDPDODATAINCONNECTOR.fun ---- *)
FUNCTION L_MC1P_FINDPDODATAINCONNECTOR : POINTER TO BYTE
VAR_INPUT
	PCONNECTOR : POINTER TO IoConfigConnector;
	UIINDEX : WORD;
	USISUBINDEX : USINT;
	XWRITEACCESS : BOOL;
END_VAR
VAR_OUTPUT
	USISIZE : USINT;
END_VAR
END_FUNCTION

(* ---- L_MC1P_GENTIMESTAMPSIMU.fun ---- *)
FUNCTION L_MC1P_GENTIMESTAMPSIMU : WORD
VAR_IN_OUT
	AXIS : AXIS_REF;
END_VAR
END_FUNCTION

(* ---- L_MC1P_GETDIGINPUTSFROMDRIVE.fun ---- *)
FUNCTION L_MC1P_GETDIGINPUTSFROMDRIVE : DWORD
VAR_IN_OUT
	AXIS : AXIS_REF;
END_VAR
END_FUNCTION

(* ---- L_MC1P_GETINSTANCENAME.fun ---- *)
FUNCTION L_MC1P_GETINSTANCENAME : STRING(L_MC1P_Constants.gc_wInstanceNchar)
VAR_INPUT
	SSTR : STRING(L_MC1P_Constants.gc_wInstanceNchar);
END_VAR
END_FUNCTION

(* ---- L_MC1P_GETIOMGRCONFIGCONNECTORLIST.fun ---- *)
FUNCTION L_MC1P_GETIOMGRCONFIGCONNECTORLIST : SysTypes.RTS_IEC_RESULT
VAR_INPUT
	PPCONNECTORLIST : POINTER TO POINTER TO IoConfigConnector;
	PNCOUNT : POINTER TO DINT;
END_VAR
END_FUNCTION

(* ---- L_MC1P_GETIOMGRCONFIGFINDCONNETOR.fun ---- *)
FUNCTION L_MC1P_GETIOMGRCONFIGFINDCONNETOR : POINTER TO IoConfigConnector
VAR_INPUT
	PCONNECTOR : POINTER TO IoConfigConnector;
END_VAR
VAR_OUTPUT
	NCOUNT : DINT := 0;
END_VAR
END_FUNCTION

(* ---- L_MC1P_GETIOMGRCONFIGFIRSTCHILD.fun ---- *)
FUNCTION L_MC1P_GETIOMGRCONFIGFIRSTCHILD : POINTER TO IoConfigConnector
VAR_INPUT
	PIOCONNECTORLIST : POINTER TO IoConfigConnector;
	PNCOUNT : POINTER TO DINT;
	PFATHER : POINTER TO IoConfigConnector;
END_VAR
END_FUNCTION

(* ---- L_MC1P_GETIOMGRCONFIGNEXTCHILD.fun ---- *)
FUNCTION L_MC1P_GETIOMGRCONFIGNEXTCHILD : POINTER TO IoConfigConnector
VAR_INPUT
	PIOCONNECTORLIST : POINTER TO IoConfigConnector;
	PNCOUNT : POINTER TO DINT;
	PFATHER : POINTER TO IoConfigConnector;
END_VAR
END_FUNCTION

(* ---- L_MC1P_GETIOMGRCONFIGPARAMETER.fun ---- *)
FUNCTION L_MC1P_GETIOMGRCONFIGPARAMETER : POINTER TO IoConfigParameter
VAR_INPUT
	PCONNECTOR : POINTER TO IoConfigConnector;
	DWPARAMETERID : DWORD;
END_VAR
END_FUNCTION

(* ---- L_MC1P_GETIOMGRCONFIGPARAMETERVALUEBYTE.fun ---- *)
FUNCTION L_MC1P_GETIOMGRCONFIGPARAMETERVALUEBYTE : BYTE
VAR_INPUT
	PPARAMETER : POINTER TO IoConfigParameter;
	PRESULT : POINTER TO UDINT;
END_VAR
END_FUNCTION

(* ---- L_MC1P_GETIOMGRCONFIGPARAMETERVALUEDWORD.fun ---- *)
FUNCTION L_MC1P_GETIOMGRCONFIGPARAMETERVALUEDWORD : DWORD
VAR_INPUT
	PPARAMETER : POINTER TO IoConfigParameter;
	PRESULT : POINTER TO UDINT;
END_VAR
END_FUNCTION

(* ---- L_MC1P_GETIOMGRCONFIGPARAMETERVALUEWORD.fun ---- *)
FUNCTION L_MC1P_GETIOMGRCONFIGPARAMETERVALUEWORD : WORD
VAR_INPUT
	PPARAMETER : POINTER TO IoConfigParameter;
	PRESULT : POINTER TO UDINT;
END_VAR
END_FUNCTION

(* ---- L_MC1P_GETRATEDTORQUEAXIS.fun ---- *)
FUNCTION L_MC1P_GETRATEDTORQUEAXIS : LREAL
VAR_IN_OUT
	AXIS : AXIS_REF;
END_VAR
END_FUNCTION

(* ---- L_MC1P_GETRATEDVELOCITYAXIS.fun ---- *)
FUNCTION L_MC1P_GETRATEDVELOCITYAXIS : LREAL
VAR_IN_OUT
	AXIS : AXIS_REF;
END_VAR
END_FUNCTION

(* ---- L_MC1P_GETTASKCYCLE.fun ---- *)
FUNCTION L_MC1P_GETTASKCYCLE : LREAL
END_FUNCTION

(* ---- L_MC1P_HLPABSDINT.fun ---- *)
FUNCTION L_MC1P_HLPABSDINT : DINT
VAR_INPUT
	DIVAR : DINT;
END_VAR
END_FUNCTION

(* ---- L_MC1P_HLPCALCPOLY5THORDERSCALED.fun ---- *)
FUNCTION L_MC1P_HLPCALCPOLY5THORDERSCALED : LREAL
VAR_OUTPUT
	LRYPOSSCALED : LREAL;
END_VAR
VAR_IN_OUT
	LRXPOSSCALED : LREAL;
	ALRKOEF : ARRAY [0..5] OF LREAL;
END_VAR
END_FUNCTION

(* ---- L_MC1P_HLPCHECKDIRECTION.fun ---- *)
FUNCTION L_MC1P_HLPCHECKDIRECTION : INT
VAR_IN_OUT
	LRPOSFIFOX : ARRAY [1..20] OF LREAL;
	LRLEN : LREAL;
END_VAR
END_FUNCTION

(* ---- L_MC1P_HLPDELTAVELTIMEEXTENDED.fun ---- *)
FUNCTION L_MC1P_HLPDELTAVELTIMEEXTENDED : BOOL
VAR_INPUT
	LRVELSTART : LREAL;
	LRACCSTART : LREAL;
	LRMAXACC : LREAL;
	LRMAXJERK : LREAL;
END_VAR
VAR_OUTPUT
	LRTIME : LREAL;
	LRDIST : LREAL;
END_VAR
END_FUNCTION

(* ---- L_MC1P_HLPFITCYCLELIM.fun ---- *)
FUNCTION L_MC1P_HLPFITCYCLELIM : BOOL
VAR_INPUT
	PLRPOS : POINTER TO LREAL;
	LRLEN : LREAL;
END_VAR
END_FUNCTION

(* ---- L_MC1P_HLPGEARRES.fun ---- *)
FUNCTION L_MC1P_HLPGEARRES : LREAL
VAR_INPUT
	LRINPUT : LREAL;
	LRNUM : LREAL;
	LRDEN : LREAL;
END_VAR
END_FUNCTION

(* ---- L_MC1P_HLPMODULOADD.fun ---- *)
FUNCTION L_MC1P_HLPMODULOADD : LREAL
VAR_INPUT
	LRINPUT : LREAL;
	LROFFSET : LREAL;
	LRLENGHT : LREAL;
END_VAR
END_FUNCTION

(* ---- L_MC1P_HLPMODULODIFF.fun ---- *)
FUNCTION L_MC1P_HLPMODULODIFF : LREAL
VAR_INPUT
	LRDIFF : LREAL;
	LRLEN : LREAL;
END_VAR
END_FUNCTION

(* ---- L_MC1P_HLPMODULOOFFSET.fun ---- *)
FUNCTION L_MC1P_HLPMODULOOFFSET : LREAL
VAR_INPUT
	LROFFSET : LREAL;
	LRLENGTH : LREAL;
	PLROFFSETBASE : POINTER TO LREAL;
END_VAR
END_FUNCTION

(* ---- L_MC1P_HLPMODULOSUB.fun ---- *)
FUNCTION L_MC1P_HLPMODULOSUB : LREAL
VAR_INPUT
	LRDIFF : LREAL;
	LRLEN : LREAL;
END_VAR
END_FUNCTION

(* ---- L_MC1P_HLPMODULOZEROPOS.fun ---- *)
FUNCTION L_MC1P_HLPMODULOZEROPOS : BOOL
VAR_INPUT
	PLRPOS : POINTER TO LREAL;
	LRLENINT : LREAL;
END_VAR
END_FUNCTION

(* ---- L_MC1P_HLPPOLY4RG.fun ---- *)
FUNCTION L_MC1P_HLPPOLY4RG : LREAL
VAR_INPUT
	LRX : LREAL;
END_VAR
END_FUNCTION

(* ---- L_MC1P_HLPPT1FILT.fun ---- *)
FUNCTION L_MC1P_HLPPT1FILT : LREAL
VAR_INPUT
	LRVALUE : LREAL;
	LRINPUT : LREAL;
	LRNEW_N : LREAL;
END_VAR
END_FUNCTION

(* ---- L_MC1P_HLPSIGNNE.fun ---- *)
FUNCTION L_MC1P_HLPSIGNNE : BOOL
VAR_INPUT
	A : LREAL;
	B : LREAL;
END_VAR
END_FUNCTION

(* ---- L_MC1P_INDEXTOPARAMETER.fun ---- *)
FUNCTION L_MC1P_INDEXTOPARAMETER : DINT
VAR_INPUT
	UIINDEX : UINT;
	USISUBINDEX : USINT;
	UIBYTELENGTH : UINT := 4;
END_VAR
END_FUNCTION

(* ---- L_MC1P_INDEXTOPARAMETER2.fun ---- *)
FUNCTION L_MC1P_INDEXTOPARAMETER2 : DINT
VAR_INPUT
	UIINDEX : UINT;
	USISUBINDEX : USINT;
	UIBYTELENGTH : UINT := 4;
	XUNSIGNED : BOOL := FALSE;
END_VAR
END_FUNCTION

(* ---- L_MC1P_LMDATAMANAGERINSERTDATA.fun ---- *)
FUNCTION L_MC1P_LMDATAMANAGERINSERTDATA : BOOL
VAR_INPUT
	ITFLMDATA : L_MC1P_ILMData;
END_VAR
END_FUNCTION

(* ---- L_MC1P_LREAL_TO_DINT.fun ---- *)
FUNCTION L_MC1P_LREAL_TO_DINT : DINT
VAR_INPUT
	LRVALUE : LREAL;
END_VAR
END_FUNCTION

(* ---- L_MC1P_LREAL_TO_DINT_TO_DWORD.fun ---- *)
FUNCTION L_MC1P_LREAL_TO_DINT_TO_DWORD : DWORD
VAR_INPUT
	LRVALUE : LREAL;
END_VAR
END_FUNCTION

(* ---- L_MC1P_LREAL_TO_DWORD.fun ---- *)
FUNCTION L_MC1P_LREAL_TO_DWORD : DWORD
VAR_INPUT
	LRVALUE : LREAL;
END_VAR
END_FUNCTION

(* ---- L_MC1P_LREAL_TO_INT.fun ---- *)
FUNCTION L_MC1P_LREAL_TO_INT : INT
VAR_INPUT
	LRVALUE : LREAL;
END_VAR
END_FUNCTION

(* ---- L_MC1P_LREAL_TO_INT_TO_WORD.fun ---- *)
FUNCTION L_MC1P_LREAL_TO_INT_TO_WORD : WORD
VAR_INPUT
	LRVALUE : LREAL;
END_VAR
END_FUNCTION

(* ---- L_MC1P_LREAL_TO_WORD.fun ---- *)
FUNCTION L_MC1P_LREAL_TO_WORD : WORD
VAR_INPUT
	LRVALUE : LREAL;
END_VAR
END_FUNCTION

(* ---- L_MC1P_LREQ.fun ---- *)
FUNCTION L_MC1P_LREQ : BOOL
VAR_INPUT
	LRVALUE : LREAL;
	LRTARGET : LREAL;
END_VAR
END_FUNCTION

(* ---- L_MC1P_LRGE.fun ---- *)
FUNCTION L_MC1P_LRGE : BOOL
VAR_INPUT
	LRVALUE : LREAL;
	LRTARGET : LREAL;
END_VAR
END_FUNCTION

(* ---- L_MC1P_LRGT.fun ---- *)
FUNCTION L_MC1P_LRGT : BOOL
VAR_INPUT
	LRVALUE : LREAL;
	LRTARGET : LREAL;
END_VAR
END_FUNCTION

(* ---- L_MC1P_LRLE.fun ---- *)
FUNCTION L_MC1P_LRLE : BOOL
VAR_INPUT
	LRVALUE : LREAL;
	LRTARGET : LREAL;
END_VAR
END_FUNCTION

(* ---- L_MC1P_LRLT.fun ---- *)
FUNCTION L_MC1P_LRLT : BOOL
VAR_INPUT
	LRVALUE : LREAL;
	LRTARGET : LREAL;
END_VAR
END_FUNCTION

(* ---- L_MC1P_LRNE.fun ---- *)
FUNCTION L_MC1P_LRNE : BOOL
VAR_INPUT
	LRVALUE : LREAL;
	LRTARGET : LREAL;
END_VAR
END_FUNCTION

(* ---- L_MC1P_MODULOCYCLE.fun ---- *)
FUNCTION L_MC1P_MODULOCYCLE : LREAL
VAR_INPUT
	LRPOSIN : LREAL;
	LRPOSITIONPERIOD : LREAL;
END_VAR
END_FUNCTION

(* ---- L_MC1P_POS_DINT_TO_LINT.fun ---- *)
FUNCTION L_MC1P_POS_DINT_TO_LINT : LINT
VAR_INPUT
	DIPOS : DINT;
	DIPOSOLD : DINT;
END_VAR
VAR_IN_OUT
	UPOS : L_MC1P_PosLINT;
END_VAR
END_FUNCTION

(* ---- L_MC1P_POSDIFFTOSPEEDINCIXXX.fun ---- *)
FUNCTION L_MC1P_POSDIFFTOSPEEDINCIXXX : DINT
VAR_INPUT
	DIPOSDIFF : DINT := 0;
	DWFACTOR : DWORD := 1000;
	DWINKPERREV : DWORD := 65536;
END_VAR
END_FUNCTION

(* ---- L_MC1P_SPEEDTOPOSDIFFINCIXXX.fun ---- *)
FUNCTION L_MC1P_SPEEDTOPOSDIFFINCIXXX : DINT
VAR_INPUT
	DISPEED : DINT := 0;
	DWFACTOR : DWORD := 1000;
	DWINKPERREV : DWORD := 65536;
END_VAR
VAR_IN_OUT
	DIRES : DINT;
END_VAR
END_FUNCTION

(* ---- L_MC1P_STVARIABLENAME_TO_DWORD.fun ---- *)
FUNCTION L_MC1P_STVARIABLENAME_TO_DWORD : BOOL
VAR_INPUT
	STVARIABLENAME : STRING;
END_VAR
VAR_OUTPUT
	DWOUT : DWORD;
END_VAR
END_FUNCTION

(* ---- L_MC1P_STVARIABLENAME_TO_INT.fun ---- *)
FUNCTION L_MC1P_STVARIABLENAME_TO_INT : BOOL
VAR_INPUT
	STVARIABLENAME : STRING;
END_VAR
VAR_OUTPUT
	IOUT : INT;
END_VAR
END_FUNCTION

(* ---- L_MC1P_STVARIABLENAME_TO_LREAL.fun ---- *)
FUNCTION L_MC1P_STVARIABLENAME_TO_LREAL : BOOL
VAR_INPUT
	STVARIABLENAME : STRING(255);
END_VAR
VAR_OUTPUT
	LROUT : LREAL;
END_VAR
END_FUNCTION

(* ---- L_MC1P_STVARIABLENAME_TO_REAL.fun ---- *)
FUNCTION L_MC1P_STVARIABLENAME_TO_REAL : BOOL
VAR_INPUT
	STVARIABLENAME : STRING;
END_VAR
VAR_OUTPUT
	ROUT : REAL;
END_VAR
END_FUNCTION

(* ---- L_MC1P_STVARIABLENAME_TO_WORD.fun ---- *)
FUNCTION L_MC1P_STVARIABLENAME_TO_WORD : BOOL
VAR_INPUT
	STVARIABLENAME : STRING;
END_VAR
VAR_OUTPUT
	WOUT : WORD;
END_VAR
END_FUNCTION

(* ---- L_MC1P_TRUNC_LINT.fun ---- *)
FUNCTION L_MC1P_TRUNC_LINT : LINT
VAR_INPUT
	LRIN : LREAL;
END_VAR
END_FUNCTION

(* ---- L_MC1P_USEHOMINGPOSITIONFROMAXISREF.fun ---- *)
FUNCTION L_MC1P_USEHOMINGPOSITIONFROMAXISREF : BOOL
VAR_INPUT
	XACTIVATE : BOOL;
END_VAR
VAR_IN_OUT
	AXIS : AXIS_REF;
END_VAR
END_FUNCTION

(* ---- L_MC1P_USEMANUALPARAMETERFROMAXISREF.fun ---- *)
FUNCTION L_MC1P_USEMANUALPARAMETERFROMAXISREF : BOOL
VAR_INPUT
	XACTIVATE : BOOL;
END_VAR
VAR_IN_OUT
	AXIS : AXIS_REF;
END_VAR
END_FUNCTION

(* ---- _AXIS_REF_9400HL.fb ---- *)
FUNCTION_BLOCK _AXIS_REF_9400HL EXTENDS _AXIS_REF_COM
VAR
	AXISEXTENSION : L_MC1P_AxisExtension_9400HL;
	MOTIONUTILS : L_MC1P_MotionUtils_9400HL;
	RETAINMANAGEMENT : L_MC1P_MotionUtilsRetainHandling;
END_VAR
END_FUNCTION_BLOCK

METHOD FB_INIT : BOOL
VAR_INPUT
	BINITRETAINS : BOOL;
	BINCOPYCODE : BOOL;
END_VAR
END_METHOD

(* ---- _AXIS_REF_9400HL_CAN.fb ---- *)
FUNCTION_BLOCK _AXIS_REF_9400HL_CAN EXTENDS _AXIS_REF_COM
VAR
	AXISEXTENSION : L_MC1P_AxisExtension_9400HL_CAN;
	MOTIONUTILS : L_MC1P_MotionUtils_9400HL_CAN;
	RETAINMANAGEMENT : L_MC1P_MotionUtilsRetainHandling;
END_VAR
END_FUNCTION_BLOCK

METHOD FB_INIT : BOOL
VAR_INPUT
	BINITRETAINS : BOOL;
	BINCOPYCODE : BOOL;
END_VAR
END_METHOD

(* ---- _AXIS_REF_COM.fb ---- *)
FUNCTION_BLOCK _AXIS_REF_COM EXTENDS _AXIS_REF_REAL
VAR
	WFATHERCONNECTORTYPE : WORD := L_MC1P_Constants.c_ConnectorTypeMotionAxisOld;
	WFATHERCONNECTORTYPE2 : WORD := L_MC1P_Constants.c_ConnectorTypeMotionAxis;
	HEVENTCOMMCYCLE : SysTypes.RTS_IEC_HANDLE := SysTypes.RTS_INVALID_HANDLE;
	HINTERFACECOMMCYCLE : SysTypes.RTS_IEC_HANDLE := SysTypes.RTS_INVALID_HANDLE;
	COMMCYCLECOUNT : DWORD;
	XCOMMERROR : BOOL;
	XCOMMWARNING : BOOL;
	WAITFORAXISDETECTION : BOOL;
END_VAR
END_FUNCTION_BLOCK

METHOD CONNECTASYNC : BOOL
END_METHOD

METHOD CALLSDODATAHANDLING
END_METHOD

METHOD CHECKCOMMUNCATION
END_METHOD

METHOD CHECKCOMMUNICATIONACYCLIC : BOOL
END_METHOD

METHOD GETMAPPEDDATA : POINTER TO BYTE
VAR_INPUT
	UIINDEX : WORD;
	USISUBINDEX : USINT;
	USISIZE : USINT;
	XWRITEACCESS : BOOL;
	PADDDATA : POINTER TO BYTE;
	PXWAITFORINITACCESS : POINTER TO BOOL;
END_VAR
VAR_OUTPUT
	EERRORID : L_IE1P_Error;
	XERROR : BOOL;
	USISIZEACT : USINT := 0;
END_VAR
END_METHOD

METHOD GETMAPPEDDATASUPPORT : BOOL
END_METHOD

METHOD HANDLESDOREADONCOMMERROR : BOOL
VAR_INPUT
	IDX : DWORD;
END_VAR
VAR_IN_OUT
	SDOREADDATA : L_DCO_SdoData;
END_VAR
END_METHOD

METHOD HANDLESDOWRITEONCOMMERROR : BOOL
VAR_INPUT
	IDX : DWORD;
END_VAR
VAR_IN_OUT
	SDOWRITEDATA : L_DCO_SdoData;
END_VAR
END_METHOD

METHOD CONFIGUREAXIS
END_METHOD

METHOD CONFIGUREAXIS2
END_METHOD

METHOD RESETAXISCONNECTOR
END_METHOD

METHOD UPDATEFATHERCONNECTOR
END_METHOD

METHOD SETAXISSIMULATION : BOOL
VAR_INPUT
	ITFAXISSIMULATION : L_MC1P_IAxisSimulationInterface;
END_VAR
END_METHOD

METHOD EVENTCALLBACK : UDINT
VAR_INPUT
	PEVENTPARAM : POINTER TO EventParam;
END_VAR
END_METHOD

METHOD REGISTEREVENT
END_METHOD

METHOD UNREGISTEREVENT
END_METHOD

METHOD GETIECADRESS
END_METHOD

(* ---- _AXIS_REF_ENC.fb ---- *)
FUNCTION_BLOCK _AXIS_REF_ENC EXTENDS _AXIS_REF_COM
VAR_INPUT
	DIENCODERPOSITION : DINT;
	XENCODERPOSVALID : BOOL := TRUE;
	POSSIGNALPROCESSING : L_MC1P_IPosSignalProcessing;
END_VAR
VAR
	WENCFILTERCYCLES : WORD := 1;
	WENCFILTERCYCLESPOS : WORD := 1;
	VELFILTER : L_MC1P_MeanValueFilter;
	ENCODERCONV : L_MC1P_EncoderConv;
	UDITOTALMEASURINGRANGE : UDINT := 4294967295;
	OPTPOSQUANT : L_MC1P_OptimizePosQuantisation;
	EXTRAPOLATION : L_MC1P_Extra_Interpolation;
	LRSETVALDELAYTIME : LREAL := 0;
	ECOMPENSATIONMODE : L_MC1P_CompensationMode := L_MC1P_CompensationMode.Off;
	XISABSOLUTEENCODER : BOOL := FALSE;
	XDRIVEENABLEDINTERN : BOOL;
	USIHOMEPOSPERMANTENTSETOLD : USINT;
	XHOMEPOSPERMANTENTSETFROMINTERN : BOOL;
	XENCODERPOSVALIDOLD : BOOL;
	XENCODERPOSVALIDINT : BOOL;
	XRESETENCODERPOSHANDLING : BOOL;
	WMICSECTICKSACT : WORD;
	WMICSECTICKSOLD : WORD;
	DIVELEXACT : DINT;
	XABSENCAVAILABLE : BOOL := FALSE;
	DWABSTIMERINFASTINPUTRESOLUTION : DWORD;
	XMANIPULATEABSCOUNTER : BOOL := FALSE;
	XCOUNTEROVERFLOW : BOOL;
	LRSCALEUNITTOPOSOLD : LREAL;
	XORIENTATIONINVACTOLD : BOOL;
	SCHOMEPARAMETER_LROFFSETPOSITIONOLD : LREAL;
	XMAXVELEXCEEDED : BOOL;
	XMAXVELEXCEEDEDOLD : BOOL;
	ITFENCODERPOSFILTER : L_MC1P_IEncoderPosFilter;
	ITFENCODERPOSFILTEROLD : L_MC1P_IEncoderPosFilter;
	ITFENCODERPOSFILTEREXTERNAL : L_MC1P_IEncoderPosFilter;
	FB_MEANPOSFILTER : L_MC1P_MeanEncoderPositionFilter;
	FB_BUTTERWORTHPOSFILTER : L_MC1P_ButterworthEncoderPosFilter;
	LRBTWFILTERTIME : LREAL;
	EENCINPUTFILTER : USINT;
	WENCFILTERCYCLESACTIVE : WORD;
	DIBTWFILTERTIME : DINT;
	EENCPOSFILTERSTATE : WORD;
	EENCVELFILTERSTATE : WORD;
	WENCODERPOSHANDLING : WORD;
	XTIMESTAMPFORPOSSUPPORTED : BOOL;
	_PTASKMAPLIST : POINTER TO IoStandard.IoConfigTaskMap;
	_NTASKMAPLISTCOUNT : DINT;
	_WMODULETYPE : UINT;
	_DWINSTANCE : UDINT;
	_CONNECTOR : POINTER TO IoConfigConnector;
	EENCODERTYPE : L_Mc1P_EncoderType;
	DIINPUTPOSOLD : DINT;
	DIACTPOSUNFILTERED : DINT;
	LRRESIDUALPOSUNFILTERED : LREAL;
	XCONFIGCHANGED : BOOL;
	DWPOSTIMESTAMP : DWORD;
	POSSIGNALPROCESSINGINT : L_MC1P_PosSignalProcessing;
	XSSIENCODER : BOOL := FALSE;
	DWENCODERUPDATETIME : DWORD;
	DIACTPOS1616 : DINT;
	XACTVELFROMPOS : BOOL;
	PDWABSOLUTECOUNTERINT : POINTER TO DWORD;
	DIACTPOSRAWOLD : DINT;
	XVELEXACTSUPPORTED : BOOL;
	CMPID_CMP_LSMCFREEENCODER : DWORD := 16#1028200D;
	ENCHOMEPOSPERMANTENTSETACTIVE : BOOL;
	GETTIMEREFVALUE : DWORD;
	HOMEPOSPERMANTENTSETACTIVE : BOOL;
	WAITFORAXISDETECTION : BOOL;
END_VAR
END_FUNCTION_BLOCK

METHOD CALCACTPOSFROMHWCOUNTER : LREAL
END_METHOD

METHOD CALCACTPOSUNFILTERED : LREAL
END_METHOD

METHOD CALCACTVALUES
END_METHOD

METHOD CALCEXTRAPOLATIONVALUES
VAR_INPUT
	LRACTPOSIN : LREAL;
	LRACTVELIN : LREAL;
	LRACTACCIN : LREAL;
	LRACTTORQUEIN : LREAL;
END_VAR
VAR_OUTPUT
	LRACTPOSOUT : LREAL;
	LRACTVELOUT : LREAL;
	LRACTACCOUT : LREAL;
	LRACTTORQUEOUT : LREAL;
END_VAR
END_METHOD

METHOD CALLRECIEVEPARAMETER
END_METHOD

METHOD CHECKPLAUSIBILITYOFACTVALUES
END_METHOD

METHOD ENCODERSIGNALHANDLING : BOOL
END_METHOD

METHOD GETACTVELOCITYEXACT : LREAL
END_METHOD

METHOD PREPAREINPUTDATA : BOOL
END_METHOD

METHOD READENCODERINPUT : BOOL
VAR_INPUT
	DINEWENCPOS : DINT;
END_VAR
END_METHOD

METHOD RESETACTPOS
END_METHOD

METHOD RESETAXISCONNECTOR
END_METHOD

METHOD RESETENCODERVALUES
END_METHOD

METHOD SETENCODERFILTERINTERFACE
VAR_INPUT
	IENCODERFILTERITF : L_MC1P_IEncoderPosFilter;
END_VAR
END_METHOD

METHOD SETHOMEPOSITION2
VAR_INPUT
	POSITION : LREAL;
	RELATIVE : BOOL;
	XRESTARTPOSITIONING : BOOL := FALSE;
	EHOMEPOSINFO : L_IE1P_Error;
END_VAR
END_METHOD

METHOD ENCNEWHOMEPOSLOADED : BOOL
VAR_INPUT
	DWCALLYCLE : DWORD;
	DWDELAY : DWORD;
END_VAR
END_METHOD

METHOD ENCRESETACTPOS
END_METHOD

METHOD ENCRESETHOMEPOS
VAR_INPUT
	ERESETINFO : L_IE1P_Error;
END_VAR
END_METHOD

METHOD ENCSETHOMEPOSITION
VAR_INPUT
	POSITION : LREAL;
	RELATIVE : BOOL;
	POSDIFF : LREAL;
	EHOMEPOSINFO : L_IE1P_Error;
END_VAR
END_METHOD

METHOD ENCSIGNALVALID : BOOL
VAR_OUTPUT
	XSIGNALVALIDOLD : BOOL;
	EENCERRORID : L_IE1P_Error;
END_VAR
END_METHOD

METHOD GETACTPOSINCR : DINT
END_METHOD

METHOD GETACTPOSINCR1616 : DINT
END_METHOD

METHOD GETACTVALUES
VAR_OUTPUT
	LRACTPOS : LREAL;
	LRACTVEL : LREAL;
	LRACTACC : LREAL;
	LRACTPOSUNFILTERED : LREAL;
	LRACTPOSROUNDS : LREAL;
END_VAR
END_METHOD

METHOD GETAXISINSTANCE : POINTER TO _AXIS_REF_REAL
END_METHOD

METHOD GETCONFIGCHANGED : BOOL
END_METHOD

METHOD GETENCODERINTERFACE : L_MC1P_IEncoderInterface
END_METHOD

METHOD GETHOMEPOSAVAILABLE : BOOL
END_METHOD

METHOD SETHOMEPOSAVAILABLE
VAR_INPUT
	XHOMEPOSAVAILABLE : BOOL;
END_VAR
END_METHOD

METHOD GETVIRTUAL : BOOL
END_METHOD

METHOD CALCSCALEFUNCTIONS
VAR_INPUT
	OFFSET : DWORD;
	INDEX : WORD;
END_VAR
END_METHOD

METHOD CALLTRANSMITPARAMETER
END_METHOD

METHOD PDCONVACTPOS : DINT
VAR_INPUT
	DIINPUT : DINT;
END_VAR
END_METHOD

METHOD PDCONVACTPOSENCCONV : DINT
VAR_INPUT
	DIINPUT : DINT;
END_VAR
END_METHOD

METHOD PDCONVACTVEL : DINT
VAR_INPUT
	DIINPUT : DINT;
END_VAR
END_METHOD

METHOD PDHANDLETIMESTAMPS : DINT
VAR_INPUT
	WMICSECTICK : WORD;
END_VAR
END_METHOD

METHOD CONFIGUREAXIS
END_METHOD

METHOD CONNECTMOTIONUTILS
VAR_INPUT
	DRIVEUTILS : L_MC1P_IDriveUtils;
	AXISEXTENSION : L_MC1P_IAxisExtension;
END_VAR
END_METHOD

METHOD CALCAFTERREADINPUTS : INT
END_METHOD

METHOD CALCBEFOREREADINPUTS : INT
END_METHOD

METHOD CALCBEFOREWRITEOUTPUTS : INT
END_METHOD

METHOD FB_INIT : BOOL
VAR_INPUT
	BINITRETAINS : BOOL;
	BINCOPYCODE : BOOL;
END_VAR
END_METHOD

METHOD IODRVUPDATEMAPPING : UDINT
VAR_INPUT
	PTASKMAPLIST : POINTER TO IoConfigTaskMap;
	NCOUNT : DINT;
END_VAR
END_METHOD

METHOD INITIALIZE : UDINT
VAR_INPUT
	WMODULETYPE : UINT;
	DWINSTANCE : UDINT;
	PCONNECTOR : POINTER TO IoConfigConnector;
END_VAR
END_METHOD

(* ---- _AXIS_REF_ENC_BPB.fb ---- *)
FUNCTION_BLOCK _AXIS_REF_ENC_BPB EXTENDS _AXIS_REF_ENC
VAR
	AXISEXTENSION : L_MC1P_AxisExtension_EncBPB;
	MOTIONUTILS : L_MC1P_MotionUtils_EncBPB;
END_VAR
END_FUNCTION_BLOCK

METHOD FB_INIT : BOOL
VAR_INPUT
	BINITRETAINS : BOOL;
	BINCOPYCODE : BOOL;
END_VAR
END_METHOD

(* ---- _AXIS_REF_ENC_FREE.fb ---- *)
FUNCTION_BLOCK _AXIS_REF_ENC_FREE EXTENDS _AXIS_REF_ENC
VAR
	AXISEXTENSION : L_MC1P_AxisExtension_EncFree;
	MOTIONUTILS : L_MC1P_MotionUtils_EncFree;
END_VAR
END_FUNCTION_BLOCK

METHOD FB_INIT : BOOL
VAR_INPUT
	BINITRETAINS : BOOL;
	BINCOPYCODE : BOOL;
END_VAR
END_METHOD

(* ---- _AXIS_REF_ENC_I500_ECAT.fb ---- *)
FUNCTION_BLOCK _AXIS_REF_ENC_I500_ECAT EXTENDS _AXIS_REF_ENC
VAR
	AXISEXTENSION : L_MC1P_AxisExtension_Enci500;
	MOTIONUTILS : L_MC1P_MotionUtils_Enci500;
END_VAR
END_FUNCTION_BLOCK

METHOD FB_INIT : BOOL
VAR_INPUT
	BINITRETAINS : BOOL;
	BINCOPYCODE : BOOL;
END_VAR
END_METHOD

(* ---- _AXIS_REF_ENC_I900.fb ---- *)
FUNCTION_BLOCK _AXIS_REF_ENC_I900 EXTENDS _AXIS_REF_ENC
END_FUNCTION_BLOCK

METHOD HLP_INITPARREF
END_METHOD

METHOD HLP_READPARAMETER : BOOL
VAR_INPUT
	PARAMETER : DINT;
	PLRVALUE : POINTER TO LREAL;
END_VAR
END_METHOD

(* ---- _AXIS_REF_ENC_I900_CIA.fb ---- *)
FUNCTION_BLOCK _AXIS_REF_ENC_I900_CIA EXTENDS _AXIS_REF_ENC_i900_Target
END_FUNCTION_BLOCK

METHOD SETDRIVECONFIG
VAR_OUTPUT
	XDONE : BOOL;
	XERROR : BOOL;
	WERRORID : WORD;
END_VAR
END_METHOD

METHOD CALCULATESCALING : BOOL
END_METHOD

METHOD FB_INIT : BOOL
VAR_INPUT
	BINITRETAINS : BOOL;
	BINCOPYCODE : BOOL;
END_VAR
END_METHOD

(* ---- _AXIS_REF_ENC_I900_ECAT.fb ---- *)
FUNCTION_BLOCK _AXIS_REF_ENC_I900_ECAT EXTENDS _AXIS_REF_ENC
VAR
	AXISEXTENSION : L_MC1P_AxisExtension_Enci900_ECAT;
	MOTIONUTILS : L_Mc1P_MotionUtils_Enci900_ECAT;
	RETAINMANAGEMENT : L_MC1P_MotionUtilsRetainHandling;
END_VAR
END_FUNCTION_BLOCK

METHOD FB_INIT : BOOL
VAR_INPUT
	BINITRETAINS : BOOL;
	BINCOPYCODE : BOOL;
END_VAR
END_METHOD

(* ---- _AXIS_REF_ENC_I900_TARGET.fb ---- *)
FUNCTION_BLOCK _AXIS_REF_ENC_I900_TARGET EXTENDS _AXIS_REF_ENC_i900
VAR
	AXISEXTENSION : L_MC1P_AxisExtension_Enci900_Target;
	MOTIONUTILS : L_MC1P_MotionUtils_Enci900_Target;
	RETAINMANAGEMENT : L_MC1P_MotionUtilsRetainHandling;
	PI900MOTIONAXIS : POINTER TO AXIS_REF;
	DWI900MOTIONAXISERRORITFID : DWORD;
	XSSIERRORBIT : BOOL;
	XSSIERRORBITOLD : BOOL;
	XSSIERRORWASSET : BOOL;
	EREACTIONSSISTATUS1 : L_IE1P_SeverityLevel;
	EREACTIONSSISTATUS1OLD : L_IE1P_SeverityLevel;
	EREACTIONSSISTATUS1ACT : L_IE1P_SeverityLevel;
END_VAR
END_FUNCTION_BLOCK

METHOD CALLRECIEVEPARAMETER
END_METHOD

METHOD CHECKSSIENCODERSTATUS : BOOL
END_METHOD

METHOD CONFIGUREAXISCONNECTOR
END_METHOD

METHOD FINDMOTIONAXIS : BOOL
END_METHOD

METHOD CALCBEFOREREADINPUTS : INT
END_METHOD

METHOD GETIECADRESS
END_METHOD

METHOD FB_INIT : BOOL
VAR_INPUT
	BINITRETAINS : BOOL;
	BINCOPYCODE : BOOL;
END_VAR
END_METHOD

(* ---- _AXIS_REF_ENC_IO_ETC.fb ---- *)
FUNCTION_BLOCK _AXIS_REF_ENC_IO_ETC EXTENDS _AXIS_REF_ENC
VAR
	AXISEXTENSION : L_MC1P_AxisExtension_EncIOEtc;
	MOTIONUTILS : L_MC1P_MotionUtils_EncIOEtc;
END_VAR
END_FUNCTION_BLOCK

METHOD INITIALIZE : UDINT
VAR_INPUT
	WMODULETYPE : UINT;
	DWINSTANCE : UDINT;
	PCONNECTOR : POINTER TO IoConfigConnector;
END_VAR
END_METHOD

METHOD FB_INIT : BOOL
VAR_INPUT
	BINITRETAINS : BOOL;
	BINCOPYCODE : BOOL;
END_VAR
END_METHOD

(* ---- _AXIS_REF_ENC_UNIVERSAL.fb ---- *)
FUNCTION_BLOCK _AXIS_REF_ENC_UNIVERSAL EXTENDS _AXIS_REF_ENC
VAR
	FBDRIVESPECIFIC : L_MC1P_DriveSpecific_Enc_Free;
	AXISEXTENSIONFACTORY : L_MC1P_UniversalEncoderFactory;
	ITFDRIVEUTILSTOCONNECT : POINTER TO L_MC1P_IDriveUtils;
	ITFAXISEXTENSION : L_MC1P_IAxisExtension;
	UITYPE : UINT := 2;
	DRIVESPECIFICBASIC : L_MC1P_IDriveSpecificImplBase;
	WAITFORAXISDETECTION : BOOL;
END_VAR
END_FUNCTION_BLOCK

METHOD CALCAFTERREADINPUTS : INT
END_METHOD

METHOD CONNECTASYNC : BOOL
END_METHOD

METHOD CREATEAXISEXTENSION : L_MC1P_IAxisExtension
VAR_INPUT
	EAXISEXTENSIONTYPE : L_MC1P_AxisExtensionTypes;
END_VAR
END_METHOD

METHOD DISCONNECTMOTIONUTILS : BOOL
VAR_INPUT
	EDISCONNECTMODE : L_IF1P_DisconnectMode;
END_VAR
END_METHOD

METHOD FINDANDCONNECTMOTIONUTILS
END_METHOD

METHOD FINDDRIVEUTILSINMOTIONCONNECTOR : BOOL
VAR_INPUT
	PECATSLAVECONNECTOR : POINTER TO IoConfigConnector;
	SUBDEVICE : UINT;
END_VAR
END_METHOD

METHOD INITIALIZE : UDINT
VAR_INPUT
	WMODULETYPE : UINT;
	DWINSTANCE : UDINT;
	PCONNECTOR : POINTER TO IoConfigConnector;
END_VAR
END_METHOD

METHOD FB_INIT : BOOL
VAR_INPUT
	BINITRETAINS : BOOL;
	BINCOPYCODE : BOOL;
END_VAR
END_METHOD

METHOD CONNECTDEVICE : UINT
VAR_INPUT
	DEVICEMODULEHANDLER : L_IMHP_IModuleHandler;
	UISUBDEVICE : UINT := 0;
	EDISCONNECTMODE : L_IF1P_DisconnectMode;
	XDISCONNECTEXISTINGCONNECTION : BOOL;
END_VAR
VAR_OUTPUT
	ITFCONNECTIONFBSTATUS : L_IF1P_IStatus;
END_VAR
END_METHOD

METHOD DISCONNECTDEVICE : UINT
VAR_INPUT
	EDISCONNECTMODE : L_IF1P_DisconnectMode;
	XBUSYBEFORE : BOOL;
END_VAR
VAR_OUTPUT
	ITFCONNECTIONFBSTATUS : L_IF1P_IStatus;
END_VAR
END_METHOD

METHOD GEFUNCTIONTINSTANCEPOINTER : POINTER TO BYTE
END_METHOD

METHOD GETCONNECTEDDEVICE : L_IMHP_IModuleHandler
VAR_OUTPUT
	UISUBDEVICE : UINT := 0;
	XVALID : BOOL;
	ITFCONNECTIONFBSTATUS : L_IF1P_IStatus;
END_VAR
END_METHOD

METHOD GETCONNECTIONDIAGNOSTIC
VAR_OUTPUT
	WUSEDBY_COMP : WORD;
	WUSEDBY_SUBCOMP : WORD;
	WACTIVEMODE : WORD;
	WSUBDEVICE : WORD;
	SCONNECTIONSOURE : STRING;
END_VAR
END_METHOD

METHOD GETITFCONNECTSTATUS
VAR_OUTPUT
	ITFCONNECTIONFBSTATUS : L_IF1P_IStatus;
END_VAR
END_METHOD

(* ---- _AXIS_REF_GENERIC.fb ---- *)
FUNCTION_BLOCK _AXIS_REF_GENERIC EXTENDS _AXIS_REF_COM
VAR
	AXISEXTENSION : L_MC1P_AxisExtension_GenericDrive;
	MOTIONUTILS : L_MC1P_MotionUtils_GenericDrive;
	RETAINMANAGEMENT : L_MC1P_MotionUtilsRetainHandling;
END_VAR
END_FUNCTION_BLOCK

METHOD SETGENERICCONFIGURATION
VAR_INPUT
	ITFGENERICCONFIG : L_MC1P_IGenericAxisConfiguration;
END_VAR
END_METHOD

METHOD FB_INIT : BOOL
VAR_INPUT
	BINITRETAINS : BOOL;
	BINCOPYCODE : BOOL;
END_VAR
END_METHOD

(* ---- _AXIS_REF_I500.fb ---- *)
FUNCTION_BLOCK _AXIS_REF_I500 EXTENDS _AXIS_REF_COM
VAR
	CONFIGAXIS : L_MC1P_Config_i500;
	FBEXTENDEDMAPPINGACCESS : L_MC1P_ExtendedMappingAccess;
	BRAKE : L_MC1P_BrakeControl;
	WNETWORDIN1 : REFERENCE TO WORD;
	WNETWORDIN2 : REFERENCE TO WORD;
	WNETWORDIN3 : REFERENCE TO WORD;
	WNETWORDIN4 : REFERENCE TO WORD;
	WNETWORDOUT1 : REFERENCE TO WORD;
	WNETWORDOUT2 : REFERENCE TO WORD;
	PXDUMMY : POINTER TO BOOL;
	XENABLEDRIVEOLD : BOOL;
	XDEACTIVATEPOSCTRLEXTENCERROR : BOOL;
	NETWORDIN1 : WORD;
	NETWORDIN2 : WORD;
	NETWORDIN3 : WORD;
	NETWORDIN4 : WORD;
	NETWORDOUT1 : WORD;
	NETWORDOUT2 : WORD;
END_VAR
END_FUNCTION_BLOCK

(* ---- _AXIS_REF_I500_CAN.fb ---- *)
FUNCTION_BLOCK _AXIS_REF_I500_CAN EXTENDS _AXIS_REF_i500
VAR
	AXISEXTENSION : L_MC1P_AxisExtension_i500_CAN;
	MOTIONUTILS : L_MC1P_MotionUtils_i500_CAN;
END_VAR
END_FUNCTION_BLOCK

METHOD FB_INIT : BOOL
VAR_INPUT
	BINITRETAINS : BOOL;
	BINCOPYCODE : BOOL;
END_VAR
END_METHOD

(* ---- _AXIS_REF_I500_ETC.fb ---- *)
FUNCTION_BLOCK _AXIS_REF_I500_ETC EXTENDS _AXIS_REF_i500
VAR
	AXISEXTENSION : L_MC1P_AxisExtension_i500_ECAT;
	MOTIONUTILS : L_MC1P_MotionUtils_i500_ECAT;
END_VAR
END_FUNCTION_BLOCK

METHOD FB_INIT : BOOL
VAR_INPUT
	BINITRETAINS : BOOL;
	BINCOPYCODE : BOOL;
END_VAR
END_METHOD

(* ---- _AXIS_REF_I700.fb ---- *)
FUNCTION_BLOCK _AXIS_REF_I700 EXTENDS _AXIS_REF_COM
VAR
	XSLOT2 : BOOL;
	AXISEXTENSION : L_MC1P_AxisExtension_i700;
	MOTIONUTILS : L_MC1P_MotionUtils_i700;
	RETAINMANAGEMENT : L_MC1P_MotionUtilsRetainHandling;
END_VAR
END_FUNCTION_BLOCK

METHOD INITIALIZE : UDINT
VAR_INPUT
	WMODULETYPE : UINT;
	DWINSTANCE : UDINT;
	PCONNECTOR : POINTER TO IoConfigConnector;
END_VAR
END_METHOD

METHOD FB_INIT : BOOL
VAR_INPUT
	BINITRETAINS : BOOL;
	BINCOPYCODE : BOOL;
END_VAR
END_METHOD

(* ---- _AXIS_REF_I700_SLOT1.fb ---- *)
FUNCTION_BLOCK _AXIS_REF_I700_SLOT1 EXTENDS _AXIS_REF_i700
END_FUNCTION_BLOCK

METHOD FB_INIT : BOOL
VAR_INPUT
	BINITRETAINS : BOOL;
	BINCOPYCODE : BOOL;
END_VAR
END_METHOD

(* ---- _AXIS_REF_I750.fb ---- *)
FUNCTION_BLOCK _AXIS_REF_I750 EXTENDS _AXIS_REF_COM
VAR
	XSLOT2 : BOOL;
	AXISEXTENSION : L_MC1P_AxisExtension_i750;
	MOTIONUTILS : L_MC1P_MotionUtils_i750;
	RETAINMANAGEMENT : L_MC1P_MotionUtilsRetainHandling;
END_VAR
END_FUNCTION_BLOCK

METHOD FB_INIT : BOOL
VAR_INPUT
	BINITRETAINS : BOOL;
	BINCOPYCODE : BOOL;
END_VAR
END_METHOD

(* ---- _AXIS_REF_I900.fb ---- *)
FUNCTION_BLOCK _AXIS_REF_I900 EXTENDS _AXIS_REF_COM
VAR
	XSLOT2 : BOOL;
	AXISEXTENSION : L_MC1P_AxisExtension_i950;
	MOTIONUTILS : L_MC1P_MotionUtils_i950;
	RETAINMANAGEMENT : L_MC1P_MotionUtilsRetainHandling;
END_VAR
END_FUNCTION_BLOCK

METHOD FB_INIT : BOOL
VAR_INPUT
	BINITRETAINS : BOOL;
	BINCOPYCODE : BOOL;
END_VAR
END_METHOD

(* ---- _AXIS_REF_I900_CIAADV.fb ---- *)
FUNCTION_BLOCK _AXIS_REF_I900_CIAADV EXTENDS _AXIS_REF_COM
VAR
	XSLOT2 : BOOL;
	AXISEXTENSION : L_MC1P_AxisExtension_i950_CiaAdv;
	MOTIONUTILS : L_MC1P_MotionUtils_i950_CiaAdv;
	RETAINMANAGEMENT : L_MC1P_MotionUtilsRetainHandling;
END_VAR
END_FUNCTION_BLOCK

METHOD FB_INIT : BOOL
VAR_INPUT
	BINITRETAINS : BOOL;
	BINCOPYCODE : BOOL;
END_VAR
END_METHOD

(* ---- _AXIS_REF_I900_DRIVE.fb ---- *)
FUNCTION_BLOCK _AXIS_REF_I900_DRIVE EXTENDS _AXIS_REF_COM
VAR
	LRHOMETORQUELIMIT : LREAL;
	LRHOMETORQUELIMITTIME : LREAL;
	EFOLLOWINGERRORREACTIONI900 : USINT;
	INTERPOLATION : L_MC1P_DelaySetValues2;
	LRSETVALDELAYTIME : LREAL := 0;
	ECOMPENSATIONMODE : L_MC1P_CompensationMode := L_MC1P_CompensationMode.Off;
	UIPOSCTRLADAPTACTIVEVALUE : UINT;
	USIPOSCTRLADAPTIONFROM0X2985 : USINT := 0;
	POSCTRLADAPTIONCURVE : L_MC1P_PosCtrlAdaptionCurve;
	DWCOMPATIBILITYFLAGS_0X2DE0_28 : DWORD;
	WAITFORAXISDETECTION : BOOL;
END_VAR
END_FUNCTION_BLOCK

METHOD GETACTIVEPOSCTRLADAPTVALUE : LREAL
END_METHOD

METHOD CONFIGUREAXISCONNECTOR
END_METHOD

METHOD CALCSCALEFUNCTIONS
VAR_INPUT
	OFFSET : DWORD;
	INDEX : WORD;
END_VAR
END_METHOD

METHOD UPDATEDRIVEOFFSETHANDLING
VAR_INPUT
	DWACTCYCLECOUNTERVALUE : DWORD;
	XRESET : BOOL;
END_VAR
END_METHOD

METHOD HLP_INITPARREF
END_METHOD

METHOD HLP_READBOOLPARAMETER : BOOL
VAR_INPUT
	PARAMETER : DINT;
	PXVALUE : POINTER TO BOOL;
END_VAR
END_METHOD

METHOD HLP_READPARAMETER : BOOL
VAR_INPUT
	PARAMETER : DINT;
	PLRVALUE : POINTER TO LREAL;
END_VAR
END_METHOD

METHOD HLP_WRITEBOOLPARAMETER : BOOL
VAR_INPUT
	PARAMETER : DINT;
	PXVALUE : POINTER TO BOOL;
END_VAR
VAR_OUTPUT
	WERRORID : WORD;
END_VAR
END_METHOD

METHOD CALCBEFOREREADINPUTS : INT
END_METHOD

METHOD CALCBEFOREWRITEOUTPUTS : INT
END_METHOD

METHOD FB_INIT : BOOL
VAR_INPUT
	BINITRETAINS : BOOL;
	BINCOPYCODE : BOOL;
END_VAR
END_METHOD

(* ---- _AXIS_REF_I900_DRIVE_CIA.fb ---- *)
FUNCTION_BLOCK _AXIS_REF_I900_DRIVE_CIA EXTENDS _AXIS_REF_i900_Drive_Target
VAR_INPUT
	XOPMODEVIACIA402INTERFACE : BOOL;
	XCONTROLVIACIAINTERFACE : BOOL;
	XSETVALUESVIAAPPLICATION : BOOL;
	CIA_CTRL_EXT : WORD;
	CIA_OPMOD_EXT : SINT;
	WLENZECTRL_EXT : WORD;
	WTPCONTROL12 : WORD;
	WTPCONTROL34 : WORD;
	XCONTROLVIACIAINTERFACEOLD : BOOL;
	XEXTSETVALUESVALID : BOOL;
	LRSETPOSITION_EXT : LREAL;
	LRSETVELOCITY_EXT : LREAL;
	LRSETTORQUE_EXT : LREAL;
	LRSETVELOCITYLIMITHIGH_EXT : LREAL;
	LRSETVELOCITYLIMITLOW_EXT : LREAL;
	LRSETVLVELOCITY_EXT : LREAL;
END_VAR
VAR_OUTPUT
	WTPSTATUS12 : WORD;
	WTPSTATUS34 : WORD;
	LRTP1_POSEDGE : LREAL;
	LRTP1_NEGEDGE : LREAL;
	DWTP1_TIMENEGEDGE : DWORD;
	DWTP1_TIMEPOSEDGE : DWORD;
	LRTP2_POSEDGE : LREAL;
	LRTP2_NEGEDGE : LREAL;
	DWTP2_TIMENEGEDGE : DWORD;
	DWTP2_TIMEPOSEDGE : DWORD;
	LRTP3_POSEDGE : LREAL;
	LRTP3_NEGEDGE : LREAL;
	DWTP3_TIMENEGEDGE : DWORD;
	DWTP3_TIMEPOSEDGE : DWORD;
	LRTP4_POSEDGE : LREAL;
	LRTP4_NEGEDGE : LREAL;
	DWTP4_TIMENEGEDGE : DWORD;
	DWTP4_TIMEPOSEDGE : DWORD;
	LRACTCONTROLEFFORT : LREAL;
END_VAR
VAR
	WPOWID : WORD;
	CIA_CTRLOLD_EXT : WORD;
	XSETVALUESVIAAPPLICATION_INT : BOOL;
	XINTTP1ACTIVE : BOOL;
	XINTTP2ACTIVE : BOOL;
	XINTTP3ACTIVE : BOOL;
	XINTTP4ACTIVE : BOOL;
	DIDRIVEREFOFFSET : DINT;
	DIDRIVEREFOFFSETABS : DINT;
	DIDRIVEREFOFFSETABSOLD : DINT;
	XDRIVELOADPOS : BOOL;
	XIGNOREDRIVEOFFSET : BOOL;
	DIDEBUGPOS : DINT;
	REFOFFSETHANDLING : L_MC1P_i900RefOffsetHandling;
	XREFOFFSETHANDLINGCALCULATED : BOOL;
	XCONFIGCHANGED : BOOL;
	XCONFIGCHANGEDENCODER : BOOL;
	X2NDFDBACTIVE : BOOL;
	X2NDFDBOBSERVATIONACTIVE : BOOL;
	LRDIRECTIONHYSTERESISDIFFOLD : LREAL;
	LRACTCONTROLEFFORTDRIVE : LREAL;
	WLENZECTRL : REFERENCE TO WORD;
	LRSPEEDCTRLINT : REFERENCE TO LREAL;
	XNEWHOMEPOSHANDLINGCIA402ADV : BOOL;
	WTEXTREFID603F : REFERENCE TO WORD;
	WLENZEEXTSTATUSWORD : REFERENCE TO WORD;
	CIA402ADVANCEDAXIS : BOOL;
	STARTPOSFORINTERNALSTOP : LREAL;
END_VAR
END_FUNCTION_BLOCK

METHOD CALCACTVALUES
END_METHOD

METHOD CALCCONTOLLER
END_METHOD

METHOD CALCDRIVEHOMEOFFSET : DINT
VAR_INPUT
	LROLDPOS : LREAL;
	LRNEWPOSPOS : LREAL;
END_VAR
END_METHOD

METHOD CHECKFOLLOWINGERROR : BOOL
END_METHOD

METHOD CHECKPLNOTVALID : BOOL
END_METHOD

METHOD CONVERTTPPOSAPP : LREAL
VAR_INPUT
	DIPOS : DINT;
END_VAR
END_METHOD

METHOD ENABLEDRIVE : BOOL
VAR_INPUT
	XENABLE : BOOL;
END_VAR
END_METHOD

METHOD GETACTDIRECTION : MC_DIRECTION
VAR_INPUT
	XCALCULATE : BOOL;
END_VAR
END_METHOD

METHOD GETDRIVESTATE : BOOL
END_METHOD

METHOD HANDLETPCONTROL
VAR_INPUT
	WTPCONTROL : WORD;
	PWCONTROL : POINTER TO WORD;
END_VAR
VAR_IN_OUT
	XTP1ACTIVE : BOOL;
	XTP2ACTIVE : BOOL;
END_VAR
END_METHOD

METHOD RESETACTPOS
END_METHOD

METHOD RESETCONFIGCHANGED
END_METHOD

METHOD SETHOMEPOSITION2
VAR_INPUT
	POSITION : LREAL;
	RELATIVE : BOOL;
	XRESTARTPOSITIONING : BOOL := FALSE;
	EHOMEPOSINFO : L_IE1P_Error;
END_VAR
END_METHOD

METHOD PDCONVACTPOS : DINT
VAR_INPUT
	DIINPUT : DINT;
END_VAR
END_METHOD

METHOD PDCONVSETPOS : DINT
VAR_INPUT
	XSETEQACTONDISABLED : BOOL;
END_VAR
END_METHOD

METHOD PDCONVTPPOS : DINT
VAR_INPUT
	DIPOS : DINT;
END_VAR
END_METHOD

METHOD SETDRIVECONFIG
VAR_OUTPUT
	XDONE : BOOL;
	XERROR : BOOL;
	WERRORID : WORD;
END_VAR
END_METHOD

METHOD CALCPOSTOUNIT : LREAL
VAR_INPUT
	DIPOSITION : DINT;
END_VAR
END_METHOD

METHOD CALCRPMTOUNIT : LREAL
VAR_INPUT
	ISPEED : INT;
END_VAR
END_METHOD

METHOD CALCSPEEDTOUNIT : LREAL
VAR_INPUT
	DISPEED : DINT;
END_VAR
END_METHOD

METHOD CALCTORQUETOUNIT : LREAL
VAR_INPUT
	ITORQUE : INT;
END_VAR
END_METHOD

METHOD CALCUNITTOPOS : DINT
VAR_INPUT
	LRPOSITION : LREAL;
END_VAR
END_METHOD

METHOD CALCUNITTORPM : INT
VAR_INPUT
	LRVELOCITY : LREAL;
END_VAR
END_METHOD

METHOD CALCUNITTOSPEED : DINT
VAR_INPUT
	LRVELOCITY : LREAL;
END_VAR
END_METHOD

METHOD CALCUNITTOTORQUE : INT
VAR_INPUT
	LRTORQUE : LREAL;
END_VAR
END_METHOD

METHOD CALCULATESCALING : BOOL
END_METHOD

METHOD RESTOREACTPOS
VAR_INPUT
	PPOSDATA : POINTER TO L_MC1P_uRetainData;
END_VAR
END_METHOD

METHOD RETAINHANDLING : BOOL
END_METHOD

METHOD STOREACTPOS
VAR_INPUT
	PPOSDATA : POINTER TO L_MC1P_uRetainData;
END_VAR
END_METHOD

METHOD STOREADDITIONALRETAINDATA
VAR_INPUT
	PDATA : POINTER TO L_MC1P_uRetainData;
END_VAR
END_METHOD

METHOD CALCBEFOREREADINPUTS : INT
END_METHOD

METHOD GETIECADRESS
END_METHOD

METHOD RECEIVEPARAMETER2
VAR_INPUT
	WPARAMETER : WORD;
	PADRESS : POINTER TO BYTE;
	WSIZE : WORD;
	PADDDATA : POINTER TO L_SI9P_IODrvMappingData;
END_VAR
END_METHOD

METHOD RECEIVEPARAMETERCALC2
VAR_IN_OUT
	DATA : ARRAY [1..L_MC1P_Constants.gc_Rec_MaxDataIndex] OF POINTER TO L_MC1P_MappedElement;
END_VAR
END_METHOD

METHOD TRANSMITPARAMETER
VAR_INPUT
	WPARAMETER : WORD;
	PADRESS : POINTER TO BYTE;
	WSIZE : WORD;
END_VAR
END_METHOD

METHOD TRANSMITPARAMETER2
VAR_INPUT
	WPARAMETER : WORD;
	PADRESS : POINTER TO BYTE;
	WSIZE : WORD;
	PADDDATA : POINTER TO L_SI9P_IODrvMappingData;
END_VAR
END_METHOD

METHOD TRANSMITPARAMETERCALC2
VAR_IN_OUT
	DATA : ARRAY [1..L_MC1P_Constants.gc_Trans_MaxDataIndex] OF POINTER TO L_MC1P_MappedElement;
END_VAR
END_METHOD

METHOD FB_INIT : BOOL
VAR_INPUT
	BINITRETAINS : BOOL;
	BINCOPYCODE : BOOL;
END_VAR
END_METHOD

(* ---- _AXIS_REF_I900_DRIVE_TARGET.fb ---- *)
FUNCTION_BLOCK _AXIS_REF_I900_DRIVE_TARGET EXTENDS _AXIS_REF_i900_Drive
VAR
	AXISEXTENSION : L_MC1P_AxisExtension_i950_Drive;
	MOTIONUTILS : L_MC1P_MotionUtils_i950_Drive;
	RETAINMANAGEMENT : L_MC1P_MotionUtilsRetainHandling;
	ADWINTERNALMAPPEDWRITEOBJECTS : ARRAY [1..c_wMaxTransElem] OF DWORD;
	HEVENTSETERRORREACTION : SysTypes.RTS_IEC_HANDLE := SysTypes.RTS_INVALID_HANDLE;
	HINTERFACESETERRORREACTION : SysTypes.RTS_IEC_HANDLE := SysTypes.RTS_INVALID_HANDLE;
	HEVENTUPDATEACTIVEERROR : SysTypes.RTS_IEC_HANDLE := SysTypes.RTS_INVALID_HANDLE;
	HINTERFACEUPDATEACTIVEERROR : SysTypes.RTS_IEC_HANDLE := SysTypes.RTS_INVALID_HANDLE;
	XINITIALREADERRORSTATUS : BOOL := FALSE;
	USIACTIVEERRORINFO : USINT := 0;
	DWLEMERRORCODE : ARRAY [0..2] OF DWORD;
	USILEMSEVERITY : ARRAY [0..2] OF USINT;
	DWPARMONITID : DWORD;
	PIPARQSPOPTION : POINTER TO INT;
	PWPARQSPOPTIONVALID : POINTER TO WORD;
	IPARQSPOPTIONOLD : INT;
	PWPARMOTORRATEDSPEED : POINTER TO WORD;
	PWPARMOTORRATEDSPEEDVALID : POINTER TO WORD;
	WPARMOTORRATEDSPEEDOLD : WORD;
	PDWPARREFTORQUE : POINTER TO DWORD;
	PWPARREFTORQUEVALID : POINTER TO WORD;
	DWPARREFTORQUEOLD : DWORD;
	PDWPARINERTIAMOTOR : POINTER TO DWORD;
	PWPARINERTIAMOTORVALID : POINTER TO WORD;
	DWPARINERTIAMOTOROLD : DWORD;
	PUSIPARMCTRLMODE : POINTER TO USINT;
	PWPARMCTRLMODEVALID : POINTER TO WORD;
	USIPARMCTRLMODEOLD : USINT;
	PDWPARMOTORRATEDCURRENT : POINTER TO DWORD;
	PWPARMOTORRATEDCURRENTVALID : POINTER TO WORD;
	DWPARMOTORRATEDCURRENTOLD : DWORD;
	PDWPARCOMPATIBILITYMODE : POINTER TO DWORD;
	PWPARCOMPATIBILITYMODEVALID : POINTER TO WORD;
	DWPARCOMPATIBILITYMODEOLD : DWORD;
	APWPARGAINADAPTSPEED : ARRAY [1..5] OF POINTER TO WORD;
	APWPARGAINADAPTSPEEDVALID : ARRAY [1..5] OF POINTER TO WORD;
	APWPARGAINADAPTOUT : ARRAY [1..5] OF POINTER TO WORD;
	APWPARGAINADAPTOUTVALID : ARRAY [1..5] OF POINTER TO WORD;
	EQUICKSTOPOPTIONACTIVE : L_MC1P_QuickStopOption := L_MC1P_QuickStopOption.StayInQSP;
END_VAR
END_FUNCTION_BLOCK

METHOD CALCDEPENDENTTORQUEVALUES
VAR_INPUT
	DWDATA : DWORD;
END_VAR
END_METHOD

METHOD GETACTIVEQUICKSTOPOPTION : L_MC1P_QuickStopOption
END_METHOD

METHOD READINITIALREADERRORSTATUS : BOOL
END_METHOD

METHOD CALLRECIEVEPARAMETER
END_METHOD

METHOD CALLTRANSMITPARAMETER
END_METHOD

METHOD CHECKMAPPEDDATAVALID : BOOL
VAR_INPUT
	PADDDATA : POINTER TO BYTE;
	PDATA : POINTER TO POINTER TO BYTE;
END_VAR
VAR_OUTPUT
	XERROR : BOOL;
	EERRORID : L_IE1P_Error;
END_VAR
END_METHOD

METHOD GETMAPPEDDATA : POINTER TO BYTE
VAR_INPUT
	UIINDEX : WORD;
	USISUBINDEX : USINT;
	USISIZE : USINT;
	XWRITEACCESS : BOOL;
	PADDDATA : POINTER TO BYTE;
	PXWAITFORINITACCESS : POINTER TO BOOL;
END_VAR
VAR_OUTPUT
	EERRORID : L_IE1P_Error;
	XERROR : BOOL;
	USISIZEACT : USINT := 0;
END_VAR
END_METHOD

METHOD GETMAPPEDDATASUPPORT : BOOL
END_METHOD

METHOD RECEIVEPARAMETER2
VAR_INPUT
	WPARAMETER : WORD;
	PADRESS : POINTER TO BYTE;
	WSIZE : WORD;
	PADDDATA : POINTER TO L_SI9P_IODrvMappingData;
END_VAR
END_METHOD

METHOD RECEIVEPARAMETERCALC2
VAR_IN_OUT
	DATA : ARRAY [1..L_MC1P_Constants.gc_Rec_MaxDataIndex] OF POINTER TO L_MC1P_MappedElement;
END_VAR
END_METHOD

METHOD RESETMAPPEDDATA
VAR_INPUT
	PADDDATA : POINTER TO BYTE;
END_VAR
END_METHOD

METHOD TRANSMITPARAMETER2
VAR_INPUT
	WPARAMETER : WORD;
	PADRESS : POINTER TO BYTE;
	WSIZE : WORD;
	PADDDATA : POINTER TO L_SI9P_IODrvMappingData;
END_VAR
END_METHOD

METHOD TRANSMITPARAMETERCALC2
VAR_IN_OUT
	DATA : ARRAY [1..L_MC1P_Constants.gc_Trans_MaxDataIndex] OF POINTER TO L_MC1P_MappedElement;
END_VAR
END_METHOD

METHOD EVENTCALLBACK : UDINT
VAR_INPUT
	PEVENTPARAM : POINTER TO EventParam;
END_VAR
END_METHOD

METHOD REGISTEREVENT
END_METHOD

METHOD UNREGISTEREVENT
END_METHOD

METHOD ITFGETACTUALERRORCODE : DWORD
VAR_OUTPUT
	ESEVERITY : WORD;
END_VAR
END_METHOD

METHOD GETIECADRESS
END_METHOD

METHOD FB_INIT : BOOL
VAR_INPUT
	BINITRETAINS : BOOL;
	BINCOPYCODE : BOOL;
END_VAR
END_METHOD
